IF NOT FRowPrepared THEN
    SelectRow();
    FCapture.Reset();
    IF NOT FPreserveResults THEN
        ResetSubjects();
    END_IF;
    CallSubjects(Enable := FALSE);
    FRowPrepared := TRUE;
ELSE
    CallSubjects(Enable := TRUE);
    CheckResults();
    FObservationReady := TRUE;
END_IF;
END_METHOD

{region 'Documentation'}
(*!
<summary>Requests fresh subject results before the next disabled call.</summary>
*)
{endregion}
METHOD PRIVATE ResetSubjects
FInRangeSubject.Reset();
FNotInRangeSubject.Reset();
END_METHOD

{region 'Documentation'}
(*!
<summary>Selects literal expectations; only named escalation rows retain preceding subject results.</summary>
*)
{endregion}
METHOD PRIVATE SelectRow
FPreserveResults := FALSE;
CASE FRow OF
    LowerEndpoint:
        FActual := ULINT#9223372036854775807;
        FLower := ULINT#9223372036854775807;
        FUpper := ULINT#9223372036854775809;
        FExpectedInRangeResult := E_Result.Passed;
        FExpectedNotInRangeResult := E_Result.Failed;
        FExpectedFindings := 1;
    Interior:
        FActual := ULINT#9223372036854775808;
        FLower := ULINT#9223372036854775807;
        FUpper := ULINT#9223372036854775809;
        FExpectedInRangeResult := E_Result.Passed;
        FExpectedNotInRangeResult := E_Result.Failed;
        FExpectedFindings := 1;
    UpperEndpoint:
        FActual := ULINT#9223372036854775809;
        FLower := ULINT#9223372036854775807;
        FUpper := ULINT#9223372036854775809;
        FExpectedInRangeResult := E_Result.Passed;
        FExpectedNotInRangeResult := E_Result.Failed;
        FExpectedFindings := 1;
    BelowRange:
        FActual := ULINT#9223372036854775806;
        FLower := ULINT#9223372036854775807;
        FUpper := ULINT#9223372036854775809;
        FExpectedInRangeResult := E_Result.Failed;
        FExpectedNotInRangeResult := E_Result.Passed;
        FExpectedFindings := 1;
    AboveRange:
        FActual := ULINT#9223372036854775810;
        FLower := ULINT#9223372036854775807;
        FUpper := ULINT#9223372036854775809;
        FExpectedInRangeResult := E_Result.Failed;
        FExpectedNotInRangeResult := E_Result.Passed;
        FExpectedFindings := 1;
    EqualBounds:
        FActual := ULINT#9223372036854775808;
        FLower := ULINT#9223372036854775808;
        FUpper := ULINT#9223372036854775808;
        FExpectedInRangeResult := E_Result.Passed;
        FExpectedNotInRangeResult := E_Result.Failed;
        FExpectedFindings := 1;
    ReversedBounds:
        FActual := ULINT#9223372036854775808;
        FLower := ULINT#9223372036854775809;
        FUpper := ULINT#9223372036854775807;
        FExpectedInRangeResult := E_Result.Error;
        FExpectedNotInRangeResult := E_Result.Error;
        FExpectedFindings := 2;
    MinimumEndpoint:
        FActual := LowestValue;
        FLower := LowestValue;
        FUpper := HighestValue;
        FExpectedInRangeResult := E_Result.Passed;
        FExpectedNotInRangeResult := E_Result.Failed;
        FExpectedFindings := 1;
    MaximumEndpoint:
        FActual := HighestValue;
        FLower := LowestValue;
        FUpper := HighestValue;
        FExpectedInRangeResult := E_Result.Passed;
        FExpectedNotInRangeResult := E_Result.Failed;
        FExpectedFindings := 1;
    FailureBeforeInvalid:
        FActual := ULINT#9223372036854775810;
        FLower := ULINT#9223372036854775807;
        FUpper := ULINT#9223372036854775809;
        FExpectedInRangeResult := E_Result.Failed;
        FExpectedNotInRangeResult := E_Result.Passed;
        FExpectedFindings := 1;
    InvalidAfterFailure:
        FActual := ULINT#9223372036854775808;
        FLower := ULINT#9223372036854775809;
        FUpper := ULINT#9223372036854775807;
        FExpectedInRangeResult := E_Result.Error;
        FExpectedNotInRangeResult := E_Result.Error;
        FExpectedFindings := 2;
        FPreserveResults := TRUE;
ELSE
    Error(Message := 'Unknown comparison test row.');
END_CASE;
END_METHOD

END_FUNCTION_BLOCK

// ---- SelfTests/TestCases/TestSuite_AssertionComparisons/Test_AssertionDurationComparisons.TcPOU
{region 'Documentation'}
(*!
<summary>Checks duration operators at millisecond boundaries and LTIME nanosecond resolution.</summary>
<description>
Named rows separate independent comparisons by a disabled reset call.
Only explicitly marked escalation rows retain the preceding subject result.
Outer Assertions latch every observation before advancing to the next row.
Intentional findings remain in the local capture; no production algorithm is copied.
</description>
*)
{endregion}
FUNCTION_BLOCK Test_AssertionDurationComparisons EXTENDS TestCaseBase
VAR
    FEqualSubject : AssertEqual_Time;
    FNotEqualSubject : AssertNotEqual_Time;
    FEarlierThanSubject : AssertEarlierThan_Time;
    FLaterThanSubject : AssertLaterThan_Time;
    FInTimespanSubject : AssertInTimespan_Time;
    FNotInTimespanSubject : AssertNotInTimespan_Time;
    FEqualLTimeSubject : AssertEqual_LTime;
    FActual : TIME;
    FReference : TIME;
    FStart : TIME;
    FEnd : TIME;
    FActualLong : LTIME;
    FReferenceLong : LTIME;
    FExpectedEqualResult : E_Result;
    FExpectedNotEqualResult : E_Result;
    FExpectedEarlierThanResult : E_Result;
    FExpectedLaterThanResult : E_Result;
    FExpectedInTimespanResult : E_Result;
    FExpectedNotInTimespanResult : E_Result;
    FExpectedEqualLTimeResult : E_Result;
    FExpectedFindings : UDINT;
    FCapture : EventBuffer;
    FEvents : ARRAY[1..CaptureLength] OF ST_Event;
    FCaptureFifo : ST_FifoStatus;
    FCaptureStatus : ST_EventBufferStatus;
    FRow : UINT;
    FRowPrepared : BOOL;
    FPreserveResults : BOOL;
    FObservationReady : BOOL;
    FChecked : BOOL;
    FSetupValid : BOOL;
END_VAR
VAR
    FEqualResult : AssertTrue;
    FEqualResultMatches : BOOL;
    FNotEqualResult : AssertTrue;
    FNotEqualResultMatches : BOOL;
    FEarlierThanResult : AssertTrue;
    FEarlierThanResultMatches : BOOL;
    FLaterThanResult : AssertTrue;
    FLaterThanResultMatches : BOOL;
    FInTimespanResult : AssertTrue;
    FInTimespanResultMatches : BOOL;
    FNotInTimespanResult : AssertTrue;
    FNotInTimespanResultMatches : BOOL;
    FEqualLTimeResult : AssertTrue;
    FEqualLTimeResultMatches : BOOL;
    FCaptureIntegrity : AssertTrue;
    FCaptureIntegrityMatches : BOOL;
END_VAR
VAR CONSTANT
    CaptureLength : UINT := 8;
    Below : UINT := 1;
    Equal : UINT := 2;
    Above : UINT := 3;
    Outside : UINT := 4;
    EqualBounds : UINT := 5;
    ReversedBounds : UINT := 6;
    LastRow : UINT := ReversedBounds;

END_VAR

SUPER^();

{region 'Documentation'}
(*!
<summary>Collects only outer checking Assertions, never intentional subject findings.</summary>
*)
{endregion}
METHOD PROTECTED AggregateResults
VAR_INPUT
    Aggregator : I_ResultAggregator; //! Borrowed result sink owned by the outer Test Case; add this test's checking Assertions without resetting or retaining the sink.
END_VAR
Aggregator.AddProvider(Provider := FEqualResult);
Aggregator.AddProvider(Provider := FNotEqualResult);
Aggregator.AddProvider(Provider := FEarlierThanResult);
Aggregator.AddProvider(Provider := FLaterThanResult);
Aggregator.AddProvider(Provider := FInTimespanResult);
Aggregator.AddProvider(Provider := FNotInTimespanResult);
Aggregator.AddProvider(Provider := FEqualLTimeResult);
Aggregator.AddProvider(Provider := FCaptureIntegrity);
END_METHOD

{region 'Documentation'}
(*!
<summary>Calls each inherited production Assertion once using the selected row.</summary>
*)
{endregion}
METHOD PRIVATE CallSubjects
VAR_INPUT
    Enable : BOOL; //! Observation-enable input forwarded to the controlled Assertion subjects for this call.
END_VAR
FEqualSubject(Enable := Enable,
    State := E_State.Running,
    IN := FActual,
    Expected := FReference);
FNotEqualSubject(Enable := Enable,
    State := E_State.Running,
    IN := FActual,
    Expected := FReference);
FEarlierThanSubject(Enable := Enable,
    State := E_State.Running,
    IN := FActual,
    Maximum := FReference);
FLaterThanSubject(Enable := Enable,
    State := E_State.Running,
    IN := FActual,
    Minimum := FReference);
FInTimespanSubject(Enable := Enable,
    State := E_State.Running,
    IN := FActual,
    StartTime := FStart,
    EndTime := FEnd);
FNotInTimespanSubject(Enable := Enable,
    State := E_State.Running,
    IN := FActual,
    StartTime := FStart,
    EndTime := FEnd);
FEqualLTimeSubject(Enable := Enable,
    State := E_State.Running,
    IN := FActualLong,
    Expected := FReferenceLong);
END_METHOD

{region 'Documentation'}
(*!
<summary>Extends base validation with subject and checking-Assertion setup.</summary>
*)
{endregion}
METHOD PROTECTED CheckInitialization : BOOL //! TRUE when the inherited initialization check and this concrete fixture check both accept the setup.
CheckInitialization := SUPER^.CheckInitialization();
IF NOT CheckInitialization THEN
    RETURN;
END_IF;

CheckInitialization := FSetupValid
    AND FEqualResult.IsInitialized
    AND FNotEqualResult.IsInitialized
    AND FEarlierThanResult.IsInitialized
    AND FLaterThanResult.IsInitialized
    AND FInTimespanResult.IsInitialized
    AND FNotInTimespanResult.IsInitialized
    AND FEqualLTimeResult.IsInitialized
    AND FCaptureIntegrity.IsInitialized;
IF NOT CheckInitialization THEN
    EventPublisher.PublishEvent(Event := CreateFrameworkEvent(Name := Name,
        ResourceName := '',
        State := State,
        Severity := E_EventSeverity.Error,
        Message := 'Comparison selftest setup failed.'));
END_IF;
END_METHOD

{region 'Documentation'}
(*!
<summary>Checks results and isolated findings against explicit expectations.</summary>
*)
{endregion}
METHOD PRIVATE CheckResults
FEqualResultMatches := FEqualSubject.Result = FExpectedEqualResult;
FNotEqualResultMatches := FNotEqualSubject.Result = FExpectedNotEqualResult;
FEarlierThanResultMatches := FEarlierThanSubject.Result = FExpectedEarlierThanResult;
FLaterThanResultMatches := FLaterThanSubject.Result = FExpectedLaterThanResult;
FInTimespanResultMatches := FInTimespanSubject.Result = FExpectedInTimespanResult;
FNotInTimespanResultMatches := FNotInTimespanSubject.Result = FExpectedNotInTimespanResult;
FEqualLTimeResultMatches := FEqualLTimeSubject.Result = FExpectedEqualLTimeResult;
FCaptureIntegrityMatches := (FCaptureStatus.SequenceId = FExpectedFindings)
    AND (FCaptureStatus.LostEventCount = 0);
END_METHOD

{region 'Documentation'}
(*!
<summary>Configures checking Assertions; subject actions remain in the test script.</summary>
*)
{endregion}
METHOD PROTECTED Configure
VAR
    Initialized : BOOL;
END_VAR
FPreparationStateCount := 0;
FTestStateCount := 1;
FEqualResult.Initialize(Parent := THIS^,
    AssertionName := 'EqualResult');
FNotEqualResult.Initialize(Parent := THIS^,
    AssertionName := 'NotEqualResult');
FEarlierThanResult.Initialize(Parent := THIS^,
    AssertionName := 'EarlierThanResult');
FLaterThanResult.Initialize(Parent := THIS^,
    AssertionName := 'LaterThanResult');
FInTimespanResult.Initialize(Parent := THIS^,
    AssertionName := 'InTimespanResult');
FNotInTimespanResult.Initialize(Parent := THIS^,
    AssertionName := 'NotInTimespanResult');
FEqualLTimeResult.Initialize(Parent := THIS^,
    AssertionName := 'EqualLTimeResult');
FCaptureIntegrity.Initialize(Parent := THIS^,
    AssertionName := 'CaptureIntegrity');
FSetupValid := FCapture.Initialize(Buffer := FEvents,
    FifoControl := FCaptureFifo,
    Status := FCaptureStatus);
FEqualSubject.BindPublisher(Publisher := FCapture);
Initialized := FEqualSubject.Initialize(Parent := THIS^,
    AssertionName := 'EqualSubject');
FSetupValid := FSetupValid AND Initialized;
FNotEqualSubject.BindPublisher(Publisher := FCapture);
Initialized := FNotEqualSubject.Initialize(Parent := THIS^,
    AssertionName := 'NotEqualSubject');
FSetupValid := FSetupValid AND Initialized;
FEarlierThanSubject.BindPublisher(Publisher := FCapture);
Initialized := FEarlierThanSubject.Initialize(Parent := THIS^,
    AssertionName := 'EarlierThanSubject');
FSetupValid := FSetupValid AND Initialized;
FLaterThanSubject.BindPublisher(Publisher := FCapture);
Initialized := FLaterThanSubject.Initialize(Parent := THIS^,
    AssertionName := 'LaterThanSubject');
FSetupValid := FSetupValid AND Initialized;
FInTimespanSubject.BindPublisher(Publisher := FCapture);
Initialized := FInTimespanSubject.Initialize(Parent := THIS^,
    AssertionName := 'InTimespanSubject');
FSetupValid := FSetupValid AND Initialized;
FNotInTimespanSubject.BindPublisher(Publisher := FCapture);
Initialized := FNotInTimespanSubject.Initialize(Parent := THIS^,
    AssertionName := 'NotInTimespanSubject');
FSetupValid := FSetupValid AND Initialized;
FEqualLTimeSubject.BindPublisher(Publisher := FCapture);
Initialized := FEqualLTimeSubject.Initialize(Parent := THIS^,
    AssertionName := 'EqualLTimeSubject');
FSetupValid := FSetupValid AND Initialized;
END_METHOD

{region 'Documentation'}
(*!
<summary>Completes abort without asynchronous resources.</summary>
*)
{endregion}
METHOD PROTECTED ProcessAbort
VAR_INPUT
    Enable : BOOL; //! Phase permission supplied by the owning Test Case; FALSE does not authorize progression, while observation may continue.
END_VAR
IF Enable THEN
    CompleteAbort();
END_IF;
END_METHOD

{region 'Documentation'}
(*!
<summary>Latches checked observations before the next script step may proceed.</summary>
*)
{endregion}
METHOD PROTECTED ProcessAssertions
VAR_INPUT
    Enable : BOOL; //! Phase permission supplied by the owning Test Case; FALSE does not authorize progression, while observation may continue.
END_VAR
VAR
    Evaluate : BOOL;
END_VAR
Evaluate := Enable AND FObservationReady;
FEqualResult(Enable := Evaluate,
    State := State,
    IN := FEqualResultMatches);
FNotEqualResult(Enable := Evaluate,
    State := State,
    IN := FNotEqualResultMatches);
FEarlierThanResult(Enable := Evaluate,
    State := State,
    IN := FEarlierThanResultMatches);
FLaterThanResult(Enable := Evaluate,
    State := State,
    IN := FLaterThanResultMatches);
FInTimespanResult(Enable := Evaluate,
    State := State,
    IN := FInTimespanResultMatches);
FNotInTimespanResult(Enable := Evaluate,
    State := State,
    IN := FNotInTimespanResultMatches);
FEqualLTimeResult(Enable := Evaluate,
    State := State,
    IN := FEqualLTimeResultMatches);
FCaptureIntegrity(Enable := Evaluate,
    State := State,
    IN := FCaptureIntegrityMatches);
IF Evaluate THEN
    FChecked := TRUE;
END_IF;
END_METHOD

{region 'Documentation'}
(*!
<summary>No Preparation phase is required.</summary>
*)
{endregion}
METHOD PROTECTED ProcessPreparations
VAR_INPUT
    // SA0033: Required hook; this test has no Preparation phase.
    {attribute 'analysis' := '-33'}
    Enable : BOOL; //! Phase permission supplied by the owning Test Case; FALSE does not authorize progression, while observation may continue.
END_VAR
END_METHOD

{region 'Documentation'}
(*!
<summary>Restarts the script and resets the checking Assertions.</summary>
*)
{endregion}
METHOD PROTECTED ProcessReset
FRow := Below;
FRowPrepared := FALSE;
FChecked := FALSE;
FObservationReady := FALSE;
FEqualResult.Reset();
FEqualResultMatches := TRUE;
FNotEqualResult.Reset();
FNotEqualResultMatches := TRUE;
FEarlierThanResult.Reset();
FEarlierThanResultMatches := TRUE;
FLaterThanResult.Reset();
FLaterThanResultMatches := TRUE;
FInTimespanResult.Reset();
FInTimespanResultMatches := TRUE;
FNotInTimespanResult.Reset();
FNotInTimespanResultMatches := TRUE;
FEqualLTimeResult.Reset();
FEqualLTimeResultMatches := TRUE;
FCaptureIntegrity.Reset();
FCaptureIntegrityMatches := TRUE;
CompleteReset();
END_METHOD

{region 'Documentation'}
(*!
<summary>Advances one bounded script step per active PLC cycle.</summary>
*)
{endregion}
METHOD PROTECTED ProcessTests
VAR_INPUT
    Enable : BOOL; //! Phase permission supplied by the owning Test Case; FALSE does not authorize progression, while observation may continue.
END_VAR
IF NOT Enable THEN
    RETURN;
END_IF;

IF FChecked THEN
    FChecked := FALSE;
    FObservationReady := FALSE;
    IF FRow = LastRow THEN
        CompleteTests();
        RETURN;
    END_IF;
    FRow := FRow + 1;
    FRowPrepared := FALSE;
END_IF;

IF NOT FRowPrepared THEN
    SelectRow();
    FCapture.Reset();
    IF NOT FPreserveResults THEN
        ResetSubjects();
    END_IF;
    CallSubjects(Enable := FALSE);
    FRowPrepared := TRUE;
ELSE
    CallSubjects(Enable := TRUE);
    CheckResults();
    FObservationReady := TRUE;
END_IF;
END_METHOD

{region 'Documentation'}
(*!
<summary>Requests fresh subject results before the next disabled call.</summary>
*)
{endregion}
METHOD PRIVATE ResetSubjects
FEqualSubject.Reset();
FNotEqualSubject.Reset();
FEarlierThanSubject.Reset();
FLaterThanSubject.Reset();
FInTimespanSubject.Reset();
FNotInTimespanSubject.Reset();
FEqualLTimeSubject.Reset();
END_METHOD

{region 'Documentation'}
(*!
<summary>Selects literal expectations; only named escalation rows retain preceding subject results.</summary>
*)
{endregion}
METHOD PRIVATE SelectRow
FPreserveResults := FALSE;
CASE FRow OF
    Below:
        FActual := T#0ms;
        FReference := T#1ms;
        FStart := T#0ms;
        FEnd := T#2ms;
        FActualLong := LTIME#0ns;
        FReferenceLong := LTIME#1ns;
        FExpectedEqualResult := E_Result.Failed;
        FExpectedNotEqualResult := E_Result.Passed;
        FExpectedEarlierThanResult := E_Result.Passed;
        FExpectedLaterThanResult := E_Result.Failed;
        FExpectedInTimespanResult := E_Result.Passed;
        FExpectedNotInTimespanResult := E_Result.Failed;
        FExpectedEqualLTimeResult := E_Result.Failed;
        FExpectedFindings := 4;
    Equal:
        FActual := T#1ms;
        FReference := T#1ms;
        FStart := T#0ms;
        FEnd := T#2ms;
        FActualLong := LTIME#1ns;
        FReferenceLong := LTIME#1ns;
        FExpectedEqualResult := E_Result.Passed;
        FExpectedNotEqualResult := E_Result.Failed;
        FExpectedEarlierThanResult := E_Result.Failed;
        FExpectedLaterThanResult := E_Result.Failed;
        FExpectedInTimespanResult := E_Result.Passed;
        FExpectedNotInTimespanResult := E_Result.Failed;
        FExpectedEqualLTimeResult := E_Result.Passed;
        FExpectedFindings := 4;
    Above:
        FActual := T#2ms;
        FReference := T#1ms;
        FStart := T#0ms;
        FEnd := T#2ms;
        FActualLong := LTIME#2ns;
        FReferenceLong := LTIME#1ns;
        FExpectedEqualResult := E_Result.Failed;
        FExpectedNotEqualResult := E_Result.Passed;
        FExpectedEarlierThanResult := E_Result.Failed;
        FExpectedLaterThanResult := E_Result.Passed;
        FExpectedInTimespanResult := E_Result.Passed;
        FExpectedNotInTimespanResult := E_Result.Failed;
        FExpectedEqualLTimeResult := E_Result.Failed;
        FExpectedFindings := 4;
    Outside:
        FActual := T#3ms;
        FReference := T#1ms;
        FStart := T#0ms;
        FEnd := T#2ms;
        FActualLong := LTIME#0ns;
        FReferenceLong := LTIME#1ns;
        FExpectedEqualResult := E_Result.Failed;
        FExpectedNotEqualResult := E_Result.Passed;
        FExpectedEarlierThanResult := E_Result.Failed;
        FExpectedLaterThanResult := E_Result.Passed;
        FExpectedInTimespanResult := E_Result.Failed;
        FExpectedNotInTimespanResult := E_Result.Passed;
        FExpectedEqualLTimeResult := E_Result.Failed;
        FExpectedFindings := 4;
    EqualBounds:
        FActual := T#1ms;
        FReference := T#1ms;
        FStart := T#1ms;
        FEnd := T#1ms;
        FActualLong := LTIME#1ns;
        FReferenceLong := LTIME#1ns;
        FExpectedEqualResult := E_Result.Passed;
        FExpectedNotEqualResult := E_Result.Failed;
        FExpectedEarlierThanResult := E_Result.Failed;
        FExpectedLaterThanResult := E_Result.Failed;
        FExpectedInTimespanResult := E_Result.Passed;
        FExpectedNotInTimespanResult := E_Result.Failed;
        FExpectedEqualLTimeResult := E_Result.Passed;
        FExpectedFindings := 4;
    ReversedBounds:
        FActual := T#1ms;
        FReference := T#1ms;
        FStart := T#2ms;
        FEnd := T#0ms;
        FActualLong := LTIME#1ns;
        FReferenceLong := LTIME#1ns;
        FExpectedEqualResult := E_Result.Passed;
        FExpectedNotEqualResult := E_Result.Failed;
        FExpectedEarlierThanResult := E_Result.Failed;
        FExpectedLaterThanResult := E_Result.Failed;
        FExpectedInTimespanResult := E_Result.Error;
        FExpectedNotInTimespanResult := E_Result.Error;
        FExpectedEqualLTimeResult := E_Result.Passed;
        FExpectedFindings := 5;
ELSE
    Error(Message := 'Unknown comparison test row.');
END_CASE;
END_METHOD

END_FUNCTION_BLOCK

// ---- Framework/Assertions/POU/BasicTypes/LTime/AssertEqual_LTime.TcPOU
{region 'Documentation'}
(*!
<summary>Checks equality with the expected LTIME value.</summary>
*)
{endregion}
FUNCTION_BLOCK AssertEqual_LTime EXTENDS AssertionBase
VAR_INPUT
    IN : LTIME; //! Actual value checked or observed by this Assertion.
    Expected : LTIME; //! Reference value for comparison with IN.
END_VAR

SUPER^();

{region 'Documentation'}
(*!
<summary>Evaluate the typed duration relation and report higher-priority errors first.</summary>
*)
{endregion}
METHOD PROTECTED Assert
VAR
    Message : STRING(GVL_Constants.MessageLength);
    ExpectedText : STRING(GVL_Constants.AssertionValueLength);
    ActualText : STRING(GVL_Constants.AssertionValueLength);
END_VAR
IF NOT EvaluationActive THEN
    RETURN;
END_IF;

IF Result = E_Result.Error THEN
    RETURN;
END_IF;

IF Result = E_Result.Failed THEN
    RETURN;
END_IF;

IF IN <> Expected THEN
    ExpectedText := LTIME_TO_STRING(Expected);
    ActualText := LTIME_TO_STRING(IN);
    Message := CONCAT('Assertion failed: values are not equal. Expected = ',
        ExpectedText);
    Message := CONCAT(Message, ', Actual = ');
    Message := CONCAT(Message, ActualText);
    Message := CONCAT(Message, '.');
    Fail(Message := Message);
    RETURN;
END_IF;

Pass();
END_METHOD

END_FUNCTION_BLOCK

// ---- SelfTests/TestCases/TestSuite_AssertionComparisons/Test_AssertionDateNormalization.TcPOU
{region 'Documentation'}
(*!
<summary>Checks calendar-day identity and range bounds despite hidden time-of-day components.</summary>
<description>
Named rows separate independent comparisons by a disabled reset call.
Only explicitly marked escalation rows retain the preceding subject result.
Outer Assertions latch every observation before advancing to the next row.
Intentional findings remain in the local capture; no production algorithm is copied.
</description>
*)
{endregion}
FUNCTION_BLOCK Test_AssertionDateNormalization EXTENDS TestCaseBase
VAR
    FEqualSubject : AssertEqual_Date;
    FInTimespanSubject : AssertInTimespan_Date;
    FNotInTimespanSubject : AssertNotInTimespan_Date;
    FActual : DATE;
    FReference : DATE;
    FStart : DATE;
    FEnd : DATE;
    FExpectedEqualResult : E_Result;
    FExpectedInTimespanResult : E_Result;
    FExpectedNotInTimespanResult : E_Result;
    FExpectedFindings : UDINT;
    FCapture : EventBuffer;
    FEvents : ARRAY[1..CaptureLength] OF ST_Event;
    FCaptureFifo : ST_FifoStatus;
    FCaptureStatus : ST_EventBufferStatus;
    FRow : UINT;
    FRowPrepared : BOOL;
    FPreserveResults : BOOL;
    FObservationReady : BOOL;
    FChecked : BOOL;
    FSetupValid : BOOL;
END_VAR
VAR
    FEqualResult : AssertTrue;
    FEqualResultMatches : BOOL;
    FInTimespanResult : AssertTrue;
    FInTimespanResultMatches : BOOL;
    FNotInTimespanResult : AssertTrue;
    FNotInTimespanResultMatches : BOOL;
    FCaptureIntegrity : AssertTrue;
    FCaptureIntegrityMatches : BOOL;
END_VAR
VAR CONSTANT
    CaptureLength : UINT := 8;
    SameDay : UINT := 1;
    NextDay : UINT := 2;
    NormalizedEqualBounds : UINT := 3;
    ReversedDays : UINT := 4;
    LastRow : UINT := ReversedDays;

END_VAR

SUPER^();

{region 'Documentation'}
(*!
<summary>Collects only outer checking Assertions, never intentional subject findings.</summary>
*)
{endregion}
METHOD PROTECTED AggregateResults
VAR_INPUT
    Aggregator : I_ResultAggregator; //! Borrowed result sink owned by the outer Test Case; add this test's checking Assertions without resetting or retaining the sink.
END_VAR
Aggregator.AddProvider(Provider := FEqualResult);
Aggregator.AddProvider(Provider := FInTimespanResult);
Aggregator.AddProvider(Provider := FNotInTimespanResult);
Aggregator.AddProvider(Provider := FCaptureIntegrity);
END_METHOD

{region 'Documentation'}
(*!
<summary>Calls each inherited production Assertion once using the selected row.</summary>
*)
{endregion}
METHOD PRIVATE CallSubjects
VAR_INPUT
    Enable : BOOL; //! Observation-enable input forwarded to the controlled Assertion subjects for this call.
END_VAR
FEqualSubject(Enable := Enable,
    State := E_State.Running,
    IN := FActual,
    Expected := FReference);
FInTimespanSubject(Enable := Enable,
    State := E_State.Running,
    IN := FActual,
    StartTime := FStart,
    EndTime := FEnd);
FNotInTimespanSubject(Enable := Enable,
    State := E_State.Running,
    IN := FActual,
    StartTime := FStart,
    EndTime := FEnd);
END_METHOD

{region 'Documentation'}
(*!
<summary>Extends base validation with subject and checking-Assertion setup.</summary>
*)
{endregion}
METHOD PROTECTED CheckInitialization : BOOL //! TRUE when the inherited initialization check and this concrete fixture check both accept the setup.
CheckInitialization := SUPER^.CheckInitialization();
IF NOT CheckInitialization THEN
    RETURN;
END_IF;

CheckInitialization := FSetupValid
    AND FEqualResult.IsInitialized
    AND FInTimespanResult.IsInitialized
    AND FNotInTimespanResult.IsInitialized
    AND FCaptureIntegrity.IsInitialized;
IF NOT CheckInitialization THEN
    EventPublisher.PublishEvent(Event := CreateFrameworkEvent(Name := Name,
        ResourceName := '',
        State := State,
        Severity := E_EventSeverity.Error,
        Message := 'Comparison selftest setup failed.'));
END_IF;
END_METHOD

{region 'Documentation'}
(*!
<summary>Checks results and isolated findings against explicit expectations.</summary>
*)
{endregion}
METHOD PRIVATE CheckResults
FEqualResultMatches := FEqualSubject.Result = FExpectedEqualResult;
FInTimespanResultMatches := FInTimespanSubject.Result = FExpectedInTimespanResult;
FNotInTimespanResultMatches := FNotInTimespanSubject.Result = FExpectedNotInTimespanResult;
FCaptureIntegrityMatches := (FCaptureStatus.SequenceId = FExpectedFindings)
    AND (FCaptureStatus.LostEventCount = 0);
END_METHOD

{region 'Documentation'}
(*!
<summary>Configures checking Assertions; subject actions remain in the test script.</summary>
*)
{endregion}
METHOD PROTECTED Configure
VAR
    Initialized : BOOL;
END_VAR
FPreparationStateCount := 0;
FTestStateCount := 1;
FEqualResult.Initialize(Parent := THIS^,
    AssertionName := 'EqualResult');
FInTimespanResult.Initialize(Parent := THIS^,
    AssertionName := 'InTimespanResult');
FNotInTimespanResult.Initialize(Parent := THIS^,
    AssertionName := 'NotInTimespanResult');
FCaptureIntegrity.Initialize(Parent := THIS^,
    AssertionName := 'CaptureIntegrity');
FSetupValid := FCapture.Initialize(Buffer := FEvents,
    FifoControl := FCaptureFifo,
    Status := FCaptureStatus);
FEqualSubject.BindPublisher(Publisher := FCapture);
Initialized := FEqualSubject.Initialize(Parent := THIS^,
    AssertionName := 'EqualSubject');
FSetupValid := FSetupValid AND Initialized;
FInTimespanSubject.BindPublisher(Publisher := FCapture);
Initialized := FInTimespanSubject.Initialize(Parent := THIS^,
    AssertionName := 'InTimespanSubject');
FSetupValid := FSetupValid AND Initialized;
FNotInTimespanSubject.BindPublisher(Publisher := FCapture);
Initialized := FNotInTimespanSubject.Initialize(Parent := THIS^,
    AssertionName := 'NotInTimespanSubject');
FSetupValid := FSetupValid AND Initialized;
END_METHOD

{region 'Documentation'}
(*!
<summary>Completes abort without asynchronous resources.</summary>
*)
{endregion}
METHOD PROTECTED ProcessAbort
VAR_INPUT
    Enable : BOOL; //! Phase permission supplied by the owning Test Case; FALSE does not authorize progression, while observation may continue.
END_VAR
IF Enable THEN
    CompleteAbort();
END_IF;
END_METHOD

{region 'Documentation'}
(*!
<summary>Latches checked observations before the next script step may proceed.</summary>
*)
{endregion}
METHOD PROTECTED ProcessAssertions
VAR_INPUT
    Enable : BOOL; //! Phase permission supplied by the owning Test Case; FALSE does not authorize progression, while observation may continue.
END_VAR
VAR
    Evaluate : BOOL;
END_VAR
Evaluate := Enable AND FObservationReady;
FEqualResult(Enable := Evaluate,
    State := State,
    IN := FEqualResultMatches);
FInTimespanResult(Enable := Evaluate,
    State := State,
    IN := FInTimespanResultMatches);
FNotInTimespanResult(Enable := Evaluate,
    State := State,
    IN := FNotInTimespanResultMatches);
FCaptureIntegrity(Enable := Evaluate,
    State := State,
    IN := FCaptureIntegrityMatches);
IF Evaluate THEN
    FChecked := TRUE;
END_IF;
END_METHOD

{region 'Documentation'}
(*!
<summary>No Preparation phase is required.</summary>
*)
{endregion}
METHOD PROTECTED ProcessPreparations
VAR_INPUT
    // SA0033: Required hook; this test has no Preparation phase.
    {attribute 'analysis' := '-33'}
    Enable : BOOL; //! Phase permission supplied by the owning Test Case; FALSE does not authorize progression, while observation may continue.
END_VAR
END_METHOD

{region 'Documentation'}
(*!
<summary>Restarts the script and resets the checking Assertions.</summary>
*)
{endregion}
METHOD PROTECTED ProcessReset
FRow := SameDay;
FRowPrepared := FALSE;
FChecked := FALSE;
FObservationReady := FALSE;
FEqualResult.Reset();
FEqualResultMatches := TRUE;
FInTimespanResult.Reset();
FInTimespanResultMatches := TRUE;
FNotInTimespanResult.Reset();
FNotInTimespanResultMatches := TRUE;
FCaptureIntegrity.Reset();
FCaptureIntegrityMatches := TRUE;
CompleteReset();
END_METHOD

{region 'Documentation'}
(*!
<summary>Advances one bounded script step per active PLC cycle.</summary>
*)
{endregion}
METHOD PROTECTED ProcessTests
VAR_INPUT
    Enable : BOOL; //! Phase permission supplied by the owning Test Case; FALSE does not authorize progression, while observation may continue.
END_VAR
IF NOT Enable THEN
    RETURN;
END_IF;

IF FChecked THEN
    FChecked := FALSE;
    FObservationReady := FALSE;
    IF FRow = LastRow THEN
        CompleteTests();
        RETURN;
    END_IF;
    FRow := FRow + 1;
    FRowPrepared := FALSE;
END_IF;

IF NOT FRowPrepared THEN
    SelectRow();
    FCapture.Reset();
    IF NOT FPreserveResults THEN
        ResetSubjects();
    END_IF;
    CallSubjects(Enable := FALSE);
    FRowPrepared := TRUE;
ELSE
    CallSubjects(Enable := TRUE);
    CheckResults();
    FObservationReady := TRUE;
END_IF;
END_METHOD

{region 'Documentation'}
(*!
<summary>Requests fresh subject results before the next disabled call.</summary>
*)
{endregion}
METHOD PRIVATE ResetSubjects
FEqualSubject.Reset();
FInTimespanSubject.Reset();
FNotInTimespanSubject.Reset();
END_METHOD

{region 'Documentation'}
(*!
<summary>Selects literal expectations; only named escalation rows retain preceding subject results.</summary>
*)
{endregion}
METHOD PRIVATE SelectRow
FPreserveResults := FALSE;
CASE FRow OF
    SameDay:
        FActual := UDINT_TO_DATE(UDINT#172799);
        FReference := UDINT_TO_DATE(UDINT#86400);
        FStart := UDINT_TO_DATE(UDINT#86400);
        FEnd := UDINT_TO_DATE(UDINT#172799);
        FExpectedEqualResult := E_Result.Passed;
        FExpectedInTimespanResult := E_Result.Passed;
        FExpectedNotInTimespanResult := E_Result.Failed;
        FExpectedFindings := 1;
    NextDay:
        FActual := UDINT_TO_DATE(UDINT#172800);
        FReference := UDINT_TO_DATE(UDINT#86400);
        FStart := UDINT_TO_DATE(UDINT#86400);
        FEnd := UDINT_TO_DATE(UDINT#172799);
        FExpectedEqualResult := E_Result.Failed;
        FExpectedInTimespanResult := E_Result.Failed;
        FExpectedNotInTimespanResult := E_Result.Passed;
        FExpectedFindings := 2;
    NormalizedEqualBounds:
        FActual := UDINT_TO_DATE(UDINT#86400);
        FReference := UDINT_TO_DATE(UDINT#172799);
        FStart := UDINT_TO_DATE(UDINT#172799);
        FEnd := UDINT_TO_DATE(UDINT#86400);
        FExpectedEqualResult := E_Result.Passed;
        FExpectedInTimespanResult := E_Result.Passed;
        FExpectedNotInTimespanResult := E_Result.Failed;
        FExpectedFindings := 1;
    ReversedDays:
        FActual := UDINT_TO_DATE(UDINT#86400);
        FReference := UDINT_TO_DATE(UDINT#86400);
        FStart := UDINT_TO_DATE(UDINT#172800);
        FEnd := UDINT_TO_DATE(UDINT#86400);
        FExpectedEqualResult := E_Result.Passed;
        FExpectedInTimespanResult := E_Result.Error;
        FExpectedNotInTimespanResult := E_Result.Error;
        FExpectedFindings := 2;
ELSE
    Error(Message := 'Unknown comparison test row.');
END_CASE;
END_METHOD

END_FUNCTION_BLOCK

// ---- Framework/Assertions/POU/BasicTypes/Date/AssertEqual_Date.TcPOU
{region 'Documentation'}
(*!
<summary>Checks equality with the expected DATE value.</summary>
<description>

Compares calendar days only; hidden time-of-day components are ignored.

</description>
*)
{endregion}
FUNCTION_BLOCK AssertEqual_Date EXTENDS AssertionBase
VAR_INPUT
    IN : DATE; //! Actual value checked or observed by this Assertion.
    Expected : DATE; //! Reference value for comparison with IN.
END_VAR

SUPER^();

{region 'Documentation'}
(*!
<summary>Evaluate the typed temporal relation and report higher-priority errors first.</summary>
*)
{endregion}
METHOD PROTECTED Assert
VAR
    Message : STRING(GVL_Constants.MessageLength);
    ExpectedText : STRING(GVL_Constants.AssertionValueLength);
    ActualText : STRING(GVL_Constants.AssertionValueLength);
END_VAR
IF NOT EvaluationActive THEN
    RETURN;
END_IF;

IF Result = E_Result.Error THEN
    RETURN;
END_IF;

IF Result = E_Result.Failed THEN
    RETURN;
END_IF;

IF DateToDayNumber(Value := IN) <> DateToDayNumber(Value := Expected) THEN
    ExpectedText := DATE_TO_STRING(Expected);
    ActualText := DATE_TO_STRING(IN);
    Message := CONCAT('Assertion failed: values are not equal. Expected = ',
        ExpectedText);
    Message := CONCAT(Message, ', Actual = ');
    Message := CONCAT(Message, ActualText);
    Message := CONCAT(Message, '.');
    Fail(Message := Message);
    RETURN;
END_IF;

Pass();
END_METHOD

END_FUNCTION_BLOCK

// ---- Framework/Assertions/POU/Utilities/DateToDayNumber.TcPOU
{region 'Documentation'}
(*!
<summary>Returns whole calendar days since 1970-01-01; ignores any time-of-day remainder.</summary>
*)
{endregion}
FUNCTION INTERNAL DateToDayNumber : UDINT //! Whole days since 1970-01-01.
VAR_INPUT
    Value : DATE; //! Calendar date; any stored time-of-day remainder is ignored.
END_VAR
VAR CONSTANT
    SecondsPerDay : UDINT := 86400;
END_VAR

DateToDayNumber := DATE_TO_UDINT(Value) / SecondsPerDay;

END_FUNCTION

// ---- Framework/Assertions/POU/BasicTypes/Date/AssertInTimespan_Date.TcPOU
{region 'Documentation'}
(*!
<summary>Check that IN is inside the inclusive StartTime..EndTime interval.</summary>
<description>

StartTime &gt; EndTime reports Error during active evaluation; equal bounds are
valid.

Compares calendar days only; hidden time-of-day components are ignored.

</description>
*)
{endregion}
FUNCTION_BLOCK AssertInTimespan_Date EXTENDS AssertionBase
VAR_INPUT
    IN : DATE; //! Actual value checked or observed by this Assertion.
    StartTime : DATE; //! Inclusive start of the time span; must not exceed EndTime.
    EndTime : DATE; //! Inclusive end of the time span; must not precede StartTime.
END_VAR

SUPER^();

{region 'Documentation'}
(*!
<summary>Evaluate the typed temporal relation and report higher-priority errors first.</summary>
*)
{endregion}
METHOD PROTECTED Assert
VAR
    Message : STRING(GVL_Constants.MessageLength);
    StartTimeText : STRING(GVL_Constants.AssertionValueLength);
    EndTimeText : STRING(GVL_Constants.AssertionValueLength);
    ActualText : STRING(GVL_Constants.AssertionValueLength);
END_VAR
IF NOT EvaluationActive THEN
    RETURN;
END_IF;

IF Result = E_Result.Error THEN
    RETURN;
END_IF;

IF DateToDayNumber(Value := StartTime) > DateToDayNumber(Value := EndTime) THEN
    StartTimeText := DATE_TO_STRING(StartTime);
    EndTimeText := DATE_TO_STRING(EndTime);
    Message := CONCAT('Assertion error: start time exceeds end time. StartTime = ',
        StartTimeText);
    Message := CONCAT(Message, ', EndTime = ');
    Message := CONCAT(Message, EndTimeText);
    Message := CONCAT(Message, '.');
    Error(Message := Message);
    RETURN;
END_IF;

IF Result = E_Result.Failed THEN
    RETURN;
END_IF;

IF (DateToDayNumber(Value := IN) < DateToDayNumber(Value := StartTime))
    OR (DateToDayNumber(Value := IN) > DateToDayNumber(Value := EndTime)) THEN
    StartTimeText := DATE_TO_STRING(StartTime);
    EndTimeText := DATE_TO_STRING(EndTime);
    ActualText := DATE_TO_STRING(IN);
    Message := CONCAT('Assertion failed: value is outside allowed timespan. StartTime = ',
        StartTimeText);
    Message := CONCAT(Message, ', EndTime = ');
    Message := CONCAT(Message, EndTimeText);
    Message := CONCAT(Message, ', Actual = ');
    Message := CONCAT(Message, ActualText);
    Message := CONCAT(Message, '.');
    Fail(Message := Message);
    RETURN;
END_IF;

Pass();
END_METHOD

END_FUNCTION_BLOCK

// ---- Framework/Assertions/POU/BasicTypes/Date/AssertNotInTimespan_Date.TcPOU
{region 'Documentation'}
(*!
<summary>Check that IN is outside the inclusive StartTime..EndTime interval.</summary>
<description>

StartTime &gt; EndTime reports Error during active evaluation; equal bounds are
valid.

Compares calendar days only; hidden time-of-day components are ignored.

</description>
*)
{endregion}
FUNCTION_BLOCK AssertNotInTimespan_Date EXTENDS AssertionBase
VAR_INPUT
    IN : DATE; //! Actual value checked or observed by this Assertion.
    StartTime : DATE; //! Inclusive start of the time span; must not exceed EndTime.
    EndTime : DATE; //! Inclusive end of the time span; must not precede StartTime.
END_VAR

SUPER^();

{region 'Documentation'}
(*!
<summary>Evaluate the typed temporal relation and report higher-priority errors first.</summary>
*)
{endregion}
METHOD PROTECTED Assert
VAR
    Message : STRING(GVL_Constants.MessageLength);
    StartTimeText : STRING(GVL_Constants.AssertionValueLength);
    EndTimeText : STRING(GVL_Constants.AssertionValueLength);
    ActualText : STRING(GVL_Constants.AssertionValueLength);
END_VAR
IF NOT EvaluationActive THEN
    RETURN;
END_IF;

IF Result = E_Result.Error THEN
    RETURN;
END_IF;

IF DateToDayNumber(Value := StartTime) > DateToDayNumber(Value := EndTime) THEN
    StartTimeText := DATE_TO_STRING(StartTime);
    EndTimeText := DATE_TO_STRING(EndTime);
    Message := CONCAT('Assertion error: start time exceeds end time. StartTime = ',
        StartTimeText);
    Message := CONCAT(Message, ', EndTime = ');
    Message := CONCAT(Message, EndTimeText);
    Message := CONCAT(Message, '.');
    Error(Message := Message);
    RETURN;
END_IF;

IF Result = E_Result.Failed THEN
    RETURN;
END_IF;

IF (DateToDayNumber(Value := IN) >= DateToDayNumber(Value := StartTime))
    AND (DateToDayNumber(Value := IN) <= DateToDayNumber(Value := EndTime)) THEN
    StartTimeText := DATE_TO_STRING(StartTime);
    EndTimeText := DATE_TO_STRING(EndTime);
    ActualText := DATE_TO_STRING(IN);
    Message := CONCAT('Assertion failed: value is inside forbidden timespan. StartTime = ',
        StartTimeText);
    Message := CONCAT(Message, ', EndTime = ');
    Message := CONCAT(Message, EndTimeText);
    Message := CONCAT(Message, ', Actual = ');
    Message := CONCAT(Message, ActualText);
    Message := CONCAT(Message, '.');
    Fail(Message := Message);
    RETURN;
END_IF;

Pass();
END_METHOD

END_FUNCTION_BLOCK

// ---- SelfTests/TestCases/TestSuite_AssertionComparisons/Test_AssertionTODDomain.TcPOU
{region 'Documentation'}
(*!
<summary>Checks all TOD inputs at midnight and the exclusive 24-hour domain limit.</summary>
<description>
Named rows separate independent comparisons by a disabled reset call.
Only explicitly marked escalation rows retain the preceding subject result.
Outer Assertions latch every observation before advancing to the next row.
Intentional findings remain in the local capture; no production algorithm is copied.
</description>
*)
{endregion}
FUNCTION_BLOCK Test_AssertionTODDomain EXTENDS TestCaseBase
VAR
    FEqualSubject : AssertEqual_TOD;
    FInTimespanSubject : AssertInTimespan_TOD;
    FNotInTimespanSubject : AssertNotInTimespan_TOD;
    FActual : TOD;
    FReference : TOD;
    FStart : TOD;
    FEnd : TOD;
    FExpectedEqualResult : E_Result;
    FExpectedInTimespanResult : E_Result;
    FExpectedNotInTimespanResult : E_Result;
    FExpectedFindings : UDINT;
    FCapture : EventBuffer;
    FEvents : ARRAY[1..CaptureLength] OF ST_Event;
    FCaptureFifo : ST_FifoStatus;
    FCaptureStatus : ST_EventBufferStatus;
    FRow : UINT;
    FRowPrepared : BOOL;
    FPreserveResults : BOOL;
    FObservationReady : BOOL;
    FChecked : BOOL;
    FSetupValid : BOOL;
END_VAR
VAR
    FEqualResult : AssertTrue;
    FEqualResultMatches : BOOL;
    FInTimespanResult : AssertTrue;
    FInTimespanResultMatches : BOOL;
    FNotInTimespanResult : AssertTrue;
    FNotInTimespanResultMatches : BOOL;
    FCaptureIntegrity : AssertTrue;
    FCaptureIntegrityMatches : BOOL;
END_VAR
VAR CONSTANT
    CaptureLength : UINT := 8;
    Midnight : UINT := 1;
    LastValidValue : UINT := 2;
    DistinctValid : UINT := 3;
    InvalidInput : UINT := 4;
    InvalidExpected : UINT := 5;
    InvalidStart : UINT := 6;
    InvalidEnd : UINT := 7;
    ReversedValidSpan : UINT := 8;
    LastRow : UINT := ReversedValidSpan;
    Zero : TOD := TOD#00:00:00;
    LastValid : TOD := TOD#23:59:59.999;
    OneDay : TOD := UDINT_TO_TOD(UDINT#86400000);
END_VAR

SUPER^();

{region 'Documentation'}
(*!
<summary>Collects only outer checking Assertions, never intentional subject findings.</summary>
*)
{endregion}
METHOD PROTECTED AggregateResults
VAR_INPUT
    Aggregator : I_ResultAggregator; //! Borrowed result sink owned by the outer Test Case; add this test's checking Assertions without resetting or retaining the sink.
END_VAR
Aggregator.AddProvider(Provider := FEqualResult);
Aggregator.AddProvider(Provider := FInTimespanResult);
Aggregator.AddProvider(Provider := FNotInTimespanResult);
Aggregator.AddProvider(Provider := FCaptureIntegrity);
END_METHOD

{region 'Documentation'}
(*!
<summary>Calls each inherited production Assertion once using the selected row.</summary>
*)
{endregion}
METHOD PRIVATE CallSubjects
VAR_INPUT
    Enable : BOOL; //! Observation-enable input forwarded to the controlled Assertion subjects for this call.
END_VAR
FEqualSubject(Enable := Enable,
    State := E_State.Running,
    IN := FActual,
    Expected := FReference);
FInTimespanSubject(Enable := Enable,
    State := E_State.Running,
    IN := FActual,
    StartTime := FStart,
    EndTime := FEnd);
FNotInTimespanSubject(Enable := Enable,
    State := E_State.Running,
    IN := FActual,
    StartTime := FStart,
    EndTime := FEnd);
END_METHOD

{region 'Documentation'}
(*!
<summary>Extends base validation with subject and checking-Assertion setup.</summary>
*)
{endregion}
METHOD PROTECTED CheckInitialization : BOOL //! TRUE when the inherited initialization check and this concrete fixture check both accept the setup.
CheckInitialization := SUPER^.CheckInitialization();
IF NOT CheckInitialization THEN
    RETURN;
END_IF;

CheckInitialization := FSetupValid
    AND FEqualResult.IsInitialized
    AND FInTimespanResult.IsInitialized
    AND FNotInTimespanResult.IsInitialized
    AND FCaptureIntegrity.IsInitialized;
IF NOT CheckInitialization THEN
    EventPublisher.PublishEvent(Event := CreateFrameworkEvent(Name := Name,
        ResourceName := '',
        State := State,
        Severity := E_EventSeverity.Error,
        Message := 'Comparison selftest setup failed.'));
END_IF;
END_METHOD

{region 'Documentation'}
(*!
<summary>Checks results and isolated findings against explicit expectations.</summary>
*)
{endregion}
METHOD PRIVATE CheckResults
FEqualResultMatches := FEqualSubject.Result = FExpectedEqualResult;
FInTimespanResultMatches := FInTimespanSubject.Result = FExpectedInTimespanResult;
FNotInTimespanResultMatches := FNotInTimespanSubject.Result = FExpectedNotInTimespanResult;
FCaptureIntegrityMatches := (FCaptureStatus.SequenceId = FExpectedFindings)
    AND (FCaptureStatus.LostEventCount = 0);
END_METHOD

{region 'Documentation'}
(*!
<summary>Configures checking Assertions; subject actions remain in the test script.</summary>
*)
{endregion}
METHOD PROTECTED Configure
VAR
    Initialized : BOOL;
END_VAR
FPreparationStateCount := 0;
FTestStateCount := 1;
FEqualResult.Initialize(Parent := THIS^,
    AssertionName := 'EqualResult');
FInTimespanResult.Initialize(Parent := THIS^,
    AssertionName := 'InTimespanResult');
FNotInTimespanResult.Initialize(Parent := THIS^,
    AssertionName := 'NotInTimespanResult');
FCaptureIntegrity.Initialize(Parent := THIS^,
    AssertionName := 'CaptureIntegrity');
FSetupValid := FCapture.Initialize(Buffer := FEvents,
    FifoControl := FCaptureFifo,
    Status := FCaptureStatus);
FEqualSubject.BindPublisher(Publisher := FCapture);
Initialized := FEqualSubject.Initialize(Parent := THIS^,
    AssertionName := 'EqualSubject');
FSetupValid := FSetupValid AND Initialized;
FInTimespanSubject.BindPublisher(Publisher := FCapture);
Initialized := FInTimespanSubject.Initialize(Parent := THIS^,
    AssertionName := 'InTimespanSubject');
FSetupValid := FSetupValid AND Initialized;
FNotInTimespanSubject.BindPublisher(Publisher := FCapture);
Initialized := FNotInTimespanSubject.Initialize(Parent := THIS^,
    AssertionName := 'NotInTimespanSubject');
FSetupValid := FSetupValid AND Initialized;
END_METHOD

{region 'Documentation'}
(*!
<summary>Completes abort without asynchronous resources.</summary>
*)
{endregion}
METHOD PROTECTED ProcessAbort
VAR_INPUT
    Enable : BOOL; //! Phase permission supplied by the owning Test Case; FALSE does not authorize progression, while observation may continue.
END_VAR
IF Enable THEN
    CompleteAbort();
END_IF;
END_METHOD

{region 'Documentation'}
(*!
<summary>Latches checked observations before the next script step may proceed.</summary>
*)
{endregion}
METHOD PROTECTED ProcessAssertions
VAR_INPUT
    Enable : BOOL; //! Phase permission supplied by the owning Test Case; FALSE does not authorize progression, while observation may continue.
END_VAR
VAR
    Evaluate : BOOL;
END_VAR
Evaluate := Enable AND FObservationReady;
FEqualResult(Enable := Evaluate,
    State := State,
    IN := FEqualResultMatches);
FInTimespanResult(Enable := Evaluate,
    State := State,
    IN := FInTimespanResultMatches);
FNotInTimespanResult(Enable := Evaluate,
    State := State,
    IN := FNotInTimespanResultMatches);
FCaptureIntegrity(Enable := Evaluate,
    State := State,
    IN := FCaptureIntegrityMatches);
IF Evaluate THEN
    FChecked := TRUE;
END_IF;
END_METHOD

{region 'Documentation'}
(*!
<summary>No Preparation phase is required.</summary>
*)
{endregion}
METHOD PROTECTED ProcessPreparations
VAR_INPUT
    // SA0033: Required hook; this test has no Preparation phase.
    {attribute 'analysis' := '-33'}
    Enable : BOOL; //! Phase permission supplied by the owning Test Case; FALSE does not authorize progression, while observation may continue.
END_VAR
END_METHOD

{region 'Documentation'}
(*!
<summary>Restarts the script and resets the checking Assertions.</summary>
*)
{endregion}
METHOD PROTECTED ProcessReset
FRow := Midnight;
FRowPrepared := FALSE;
FChecked := FALSE;
FObservationReady := FALSE;
FEqualResult.Reset();
FEqualResultMatches := TRUE;
FInTimespanResult.Reset();
FInTimespanResultMatches := TRUE;
FNotInTimespanResult.Reset();
FNotInTimespanResultMatches := TRUE;
FCaptureIntegrity.Reset();
FCaptureIntegrityMatches := TRUE;
CompleteReset();
END_METHOD

{region 'Documentation'}
(*!
<summary>Advances one bounded script step per active PLC cycle.</summary>
*)
{endregion}
METHOD PROTECTED ProcessTests
VAR_INPUT
    Enable : BOOL; //! Phase permission supplied by the owning Test Case; FALSE does not authorize progression, while observation may continue.
END_VAR
IF NOT Enable THEN
    RETURN;
END_IF;

IF FChecked THEN
    FChecked := FALSE;
    FObservationReady := FALSE;
    IF FRow = LastRow THEN
        CompleteTests();
        RETURN;
    END_IF;
    FRow := FRow + 1;
    FRowPrepared := FALSE;
END_IF;

IF NOT FRowPrepared THEN
    SelectRow();
    FCapture.Reset();
    IF NOT FPreserveResults THEN
        ResetSubjects();
    END_IF;
    CallSubjects(Enable := FALSE);
    FRowPrepared := TRUE;
ELSE
    CallSubjects(Enable := TRUE);
    CheckResults();
    FObservationReady := TRUE;
END_IF;
END_METHOD

{region 'Documentation'}
(*!
<summary>Requests fresh subject results before the next disabled call.</summary>
*)
{endregion}
METHOD PRIVATE ResetSubjects
FEqualSubject.Reset();
FInTimespanSubject.Reset();
FNotInTimespanSubject.Reset();
END_METHOD

{region 'Documentation'}
(*!
<summary>Selects literal expectations; only named escalation rows retain preceding subject results.</summary>
*)
{endregion}
METHOD PRIVATE SelectRow
FPreserveResults := FALSE;
CASE FRow OF
    Midnight:
        FActual := Zero;
        FReference := Zero;
        FStart := Zero;
        FEnd := LastValid;
        FExpectedEqualResult := E_Result.Passed;
        FExpectedInTimespanResult := E_Result.Passed;
        FExpectedNotInTimespanResult := E_Result.Failed;
        FExpectedFindings := 1;
    LastValidValue:
        FActual := LastValid;
        FReference := LastValid;
        FStart := Zero;
        FEnd := LastValid;
        FExpectedEqualResult := E_Result.Passed;
        FExpectedInTimespanResult := E_Result.Passed;
        FExpectedNotInTimespanResult := E_Result.Failed;
        FExpectedFindings := 1;
    DistinctValid:
        FActual := Zero;
        FReference := LastValid;
        FStart := Zero;
        FEnd := LastValid;
        FExpectedEqualResult := E_Result.Failed;
        FExpectedInTimespanResult := E_Result.Passed;
        FExpectedNotInTimespanResult := E_Result.Failed;
        FExpectedFindings := 2;
    InvalidInput:
        FActual := OneDay;
        FReference := Zero;
        FStart := Zero;
        FEnd := LastValid;
        FExpectedEqualResult := E_Result.Error;
        FExpectedInTimespanResult := E_Result.Error;
        FExpectedNotInTimespanResult := E_Result.Error;
        FExpectedFindings := 3;
    InvalidExpected:
        FActual := Zero;
        FReference := OneDay;
        FStart := Zero;
        FEnd := LastValid;
        FExpectedEqualResult := E_Result.Error;
        FExpectedInTimespanResult := E_Result.Passed;
        FExpectedNotInTimespanResult := E_Result.Failed;
        FExpectedFindings := 2;
    InvalidStart:
        FActual := Zero;
        FReference := Zero;
        FStart := OneDay;
        FEnd := LastValid;
        FExpectedEqualResult := E_Result.Passed;
        FExpectedInTimespanResult := E_Result.Error;
        FExpectedNotInTimespanResult := E_Result.Error;
        FExpectedFindings := 2;
    InvalidEnd:
        FActual := Zero;
        FReference := Zero;
        FStart := Zero;
        FEnd := OneDay;
        FExpectedEqualResult := E_Result.Passed;
        FExpectedInTimespanResult := E_Result.Error;
        FExpectedNotInTimespanResult := E_Result.Error;
        FExpectedFindings := 2;
    ReversedValidSpan:
        FActual := Zero;
        FReference := Zero;
        FStart := LastValid;
        FEnd := Zero;
        FExpectedEqualResult := E_Result.Passed;
        FExpectedInTimespanResult := E_Result.Error;
        FExpectedNotInTimespanResult := E_Result.Error;
        FExpectedFindings := 2;
ELSE
    Error(Message := 'Unknown comparison test row.');
END_CASE;
END_METHOD

END_FUNCTION_BLOCK

// ---- SelfTests/TestCases/TestSuite_AssertionComparisons/Test_AssertionLTODDomain.TcPOU
{region 'Documentation'}
(*!
<summary>Checks all LTOD inputs at midnight and the exclusive 24-hour domain limit.</summary>
<description>
Named rows separate independent comparisons by a disabled reset call.
Only explicitly marked escalation rows retain the preceding subject result.
Outer Assertions latch every observation before advancing to the next row.
Intentional findings remain in the local capture; no production algorithm is copied.
</description>
*)
{endregion}
FUNCTION_BLOCK Test_AssertionLTODDomain EXTENDS TestCaseBase
VAR
    FEqualSubject : AssertEqual_LTOD;
    FInTimespanSubject : AssertInTimespan_LTOD;
    FNotInTimespanSubject : AssertNotInTimespan_LTOD;
    FActual : LTOD;
    FReference : LTOD;
    FStart : LTOD;
    FEnd : LTOD;
    FExpectedEqualResult : E_Result;
    FExpectedInTimespanResult : E_Result;
    FExpectedNotInTimespanResult : E_Result;
    FExpectedFindings : UDINT;
    FCapture : EventBuffer;
    FEvents : ARRAY[1..CaptureLength] OF ST_Event;
    FCaptureFifo : ST_FifoStatus;
    FCaptureStatus : ST_EventBufferStatus;
    FRow : UINT;
    FRowPrepared : BOOL;
    FPreserveResults : BOOL;
    FObservationReady : BOOL;
    FChecked : BOOL;
    FSetupValid : BOOL;
END_VAR
VAR
    FEqualResult : AssertTrue;
    FEqualResultMatches : BOOL;
    FInTimespanResult : AssertTrue;
    FInTimespanResultMatches : BOOL;
    FNotInTimespanResult : AssertTrue;
    FNotInTimespanResultMatches : BOOL;
    FCaptureIntegrity : AssertTrue;
    FCaptureIntegrityMatches : BOOL;
END_VAR
VAR CONSTANT
    CaptureLength : UINT := 8;
    Midnight : UINT := 1;
    LastValidValue : UINT := 2;
    DistinctValid : UINT := 3;
    InvalidInput : UINT := 4;
    InvalidExpected : UINT := 5;
    InvalidStart : UINT := 6;
    InvalidEnd : UINT := 7;
    ReversedValidSpan : UINT := 8;
    LastRow : UINT := ReversedValidSpan;
    Zero : LTOD := LTOD#00:00:00;
    LastValid : LTOD := LTOD#23:59:59.999999999;
    OneDay : LTOD := ULINT_TO_LTOD(ULINT#86400000000000);
END_VAR

SUPER^();

{region 'Documentation'}
(*!
<summary>Collects only outer checking Assertions, never intentional subject findings.</summary>
*)
{endregion}
METHOD PROTECTED AggregateResults
VAR_INPUT
    Aggregator : I_ResultAggregator; //! Borrowed result sink owned by the outer Test Case; add this test's checking Assertions without resetting or retaining the sink.
END_VAR
Aggregator.AddProvider(Provider := FEqualResult);
Aggregator.AddProvider(Provider := FInTimespanResult);
Aggregator.AddProvider(Provider := FNotInTimespanResult);
Aggregator.AddProvider(Provider := FCaptureIntegrity);
END_METHOD

{region 'Documentation'}
(*!
<summary>Calls each inherited production Assertion once using the selected row.</summary>
*)
{endregion}
METHOD PRIVATE CallSubjects
VAR_INPUT
    Enable : BOOL; //! Observation-enable input forwarded to the controlled Assertion subjects for this call.
END_VAR
FEqualSubject(Enable := Enable,
    State := E_State.Running,
    IN := FActual,
    Expected := FReference);
FInTimespanSubject(Enable := Enable,
    State := E_State.Running,
    IN := FActual,
    StartTime := FStart,
    EndTime := FEnd);
FNotInTimespanSubject(Enable := Enable,
    State := E_State.Running,
    IN := FActual,
    StartTime := FStart,
    EndTime := FEnd);
END_METHOD

{region 'Documentation'}
(*!
<summary>Extends base validation with subject and checking-Assertion setup.</summary>
*)
{endregion}
METHOD PROTECTED CheckInitialization : BOOL //! TRUE when the inherited initialization check and this concrete fixture check both accept the setup.
CheckInitialization := SUPER^.CheckInitialization();
IF NOT CheckInitialization THEN
    RETURN;
END_IF;

CheckInitialization := FSetupValid
    AND FEqualResult.IsInitialized
    AND FInTimespanResult.IsInitialized
    AND FNotInTimespanResult.IsInitialized
    AND FCaptureIntegrity.IsInitialized;
IF NOT CheckInitialization THEN
    EventPublisher.PublishEvent(Event := CreateFrameworkEvent(Name := Name,
        ResourceName := '',
        State := State,
        Severity := E_EventSeverity.Error,
        Message := 'Comparison selftest setup failed.'));
END_IF;
END_METHOD

{region 'Documentation'}
(*!
<summary>Checks results and isolated findings against explicit expectations.</summary>
*)
{endregion}
METHOD PRIVATE CheckResults
FEqualResultMatches := FEqualSubject.Result = FExpectedEqualResult;
FInTimespanResultMatches := FInTimespanSubject.Result = FExpectedInTimespanResult;
FNotInTimespanResultMatches := FNotInTimespanSubject.Result = FExpectedNotInTimespanResult;
FCaptureIntegrityMatches := (FCaptureStatus.SequenceId = FExpectedFindings)
    AND (FCaptureStatus.LostEventCount = 0);
END_METHOD

{region 'Documentation'}
(*!
<summary>Configures checking Assertions; subject actions remain in the test script.</summary>
*)
{endregion}
METHOD PROTECTED Configure
VAR
    Initialized : BOOL;
END_VAR
FPreparationStateCount := 0;
FTestStateCount := 1;
FEqualResult.Initialize(Parent := THIS^,
    AssertionName := 'EqualResult');
FInTimespanResult.Initialize(Parent := THIS^,
    AssertionName := 'InTimespanResult');
FNotInTimespanResult.Initialize(Parent := THIS^,
    AssertionName := 'NotInTimespanResult');
FCaptureIntegrity.Initialize(Parent := THIS^,
    AssertionName := 'CaptureIntegrity');
FSetupValid := FCapture.Initialize(Buffer := FEvents,
    FifoControl := FCaptureFifo,
    Status := FCaptureStatus);
FEqualSubject.BindPublisher(Publisher := FCapture);
Initialized := FEqualSubject.Initialize(Parent := THIS^,
    AssertionName := 'EqualSubject');
FSetupValid := FSetupValid AND Initialized;
FInTimespanSubject.BindPublisher(Publisher := FCapture);
Initialized := FInTimespanSubject.Initialize(Parent := THIS^,
    AssertionName := 'InTimespanSubject');
FSetupValid := FSetupValid AND Initialized;
FNotInTimespanSubject.BindPublisher(Publisher := FCapture);
Initialized := FNotInTimespanSubject.Initialize(Parent := THIS^,
    AssertionName := 'NotInTimespanSubject');
FSetupValid := FSetupValid AND Initialized;
END_METHOD

{region 'Documentation'}
(*!
<summary>Completes abort without asynchronous resources.</summary>
*)
{endregion}
METHOD PROTECTED ProcessAbort
VAR_INPUT
    Enable : BOOL; //! Phase permission supplied by the owning Test Case; FALSE does not authorize progression, while observation may continue.
END_VAR
IF Enable THEN
    CompleteAbort();
END_IF;
END_METHOD

{region 'Documentation'}
(*!
<summary>Latches checked observations before the next script step may proceed.</summary>
*)
{endregion}
METHOD PROTECTED ProcessAssertions
VAR_INPUT
    Enable : BOOL; //! Phase permission supplied by the owning Test Case; FALSE does not authorize progression, while observation may continue.
END_VAR
VAR
    Evaluate : BOOL;
END_VAR
Evaluate := Enable AND FObservationReady;
FEqualResult(Enable := Evaluate,
    State := State,
    IN := FEqualResultMatches);
FInTimespanResult(Enable := Evaluate,
    State := State,
    IN := FInTimespanResultMatches);
FNotInTimespanResult(Enable := Evaluate,
    State := State,
    IN := FNotInTimespanResultMatches);
FCaptureIntegrity(Enable := Evaluate,
    State := State,
    IN := FCaptureIntegrityMatches);
IF Evaluate THEN
    FChecked := TRUE;
END_IF;
END_METHOD

{region 'Documentation'}
(*!
<summary>No Preparation phase is required.</summary>
*)
{endregion}
METHOD PROTECTED ProcessPreparations
VAR_INPUT
    // SA0033: Required hook; this test has no Preparation phase.
    {attribute 'analysis' := '-33'}
    Enable : BOOL; //! Phase permission supplied by the owning Test Case; FALSE does not authorize progression, while observation may continue.
END_VAR
END_METHOD

{region 'Documentation'}
(*!
<summary>Restarts the script and resets the checking Assertions.</summary>
*)
{endregion}
METHOD PROTECTED ProcessReset
FRow := Midnight;
FRowPrepared := FALSE;
FChecked := FALSE;
FObservationReady := FALSE;
FEqualResult.Reset();
FEqualResultMatches := TRUE;
FInTimespanResult.Reset();
FInTimespanResultMatches := TRUE;
FNotInTimespanResult.Reset();
FNotInTimespanResultMatches := TRUE;
FCaptureIntegrity.Reset();
FCaptureIntegrityMatches := TRUE;
CompleteReset();
END_METHOD

{region 'Documentation'}
(*!
<summary>Advances one bounded script step per active PLC cycle.</summary>
*)
{endregion}
METHOD PROTECTED ProcessTests
VAR_INPUT
    Enable : BOOL; //! Phase permission supplied by the owning Test Case; FALSE does not authorize progression, while observation may continue.
END_VAR
IF NOT Enable THEN
    RETURN;
END_IF;

IF FChecked THEN
    FChecked := FALSE;
    FObservationReady := FALSE;
    IF FRow = LastRow THEN
        CompleteTests();
        RETURN;
    END_IF;
    FRow := FRow + 1;
    FRowPrepared := FALSE;
END_IF;

IF NOT FRowPrepared THEN
    SelectRow();
    FCapture.Reset();
    IF NOT FPreserveResults THEN
        ResetSubjects();
    END_IF;
    CallSubjects(Enable := FALSE);
    FRowPrepared := TRUE;
ELSE
    CallSubjects(Enable := TRUE);
    CheckResults();
    FObservationReady := TRUE;
END_IF;
END_METHOD

{region 'Documentation'}
(*!
<summary>Requests fresh subject results before the next disabled call.</summary>
*)
{endregion}
METHOD PRIVATE ResetSubjects
FEqualSubject.Reset();
FInTimespanSubject.Reset();
FNotInTimespanSubject.Reset();
END_METHOD

{region 'Documentation'}
(*!
<summary>Selects literal expectations; only named escalation rows retain preceding subject results.</summary>
*)
{endregion}
METHOD PRIVATE SelectRow
FPreserveResults := FALSE;
CASE FRow OF
    Midnight:
        FActual := Zero;
        FReference := Zero;
        FStart := Zero;
        FEnd := LastValid;
        FExpectedEqualResult := E_Result.Passed;
        FExpectedInTimespanResult := E_Result.Passed;
        FExpectedNotInTimespanResult := E_Result.Failed;
        FExpectedFindings := 1;
    LastValidValue:
        FActual := LastValid;
        FReference := LastValid;
        FStart := Zero;
        FEnd := LastValid;
        FExpectedEqualResult := E_Result.Passed;
        FExpectedInTimespanResult := E_Result.Passed;
        FExpectedNotInTimespanResult := E_Result.Failed;
        FExpectedFindings := 1;
    DistinctValid:
        FActual := Zero;
        FReference := LastValid;
        FStart := Zero;
        FEnd := LastValid;
        FExpectedEqualResult := E_Result.Failed;
        FExpectedInTimespanResult := E_Result.Passed;
        FExpectedNotInTimespanResult := E_Result.Failed;
        FExpectedFindings := 2;
    InvalidInput:
        FActual := OneDay;
        FReference := Zero;
        FStart := Zero;
        FEnd := LastValid;
        FExpectedEqualResult := E_Result.Error;
        FExpectedInTimespanResult := E_Result.Error;
        FExpectedNotInTimespanResult := E_Result.Error;
        FExpectedFindings := 3;
    InvalidExpected:
        FActual := Zero;
        FReference := OneDay;
        FStart := Zero;
        FEnd := LastValid;
        FExpectedEqualResult := E_Result.Error;
        FExpectedInTimespanResult := E_Result.Passed;
        FExpectedNotInTimespanResult := E_Result.Failed;
        FExpectedFindings := 2;
    InvalidStart:
        FActual := Zero;
        FReference := Zero;
        FStart := OneDay;
        FEnd := LastValid;
        FExpectedEqualResult := E_Result.Passed;
        FExpectedInTimespanResult := E_Result.Error;
        FExpectedNotInTimespanResult := E_Result.Error;
        FExpectedFindings := 2;
    InvalidEnd:
        FActual := Zero;
        FReference := Zero;
        FStart := Zero;
        FEnd := OneDay;
        FExpectedEqualResult := E_Result.Passed;
        FExpectedInTimespanResult := E_Result.Error;
        FExpectedNotInTimespanResult := E_Result.Error;
        FExpectedFindings := 2;
    ReversedValidSpan:
        FActual := Zero;
        FReference := Zero;
        FStart := LastValid;
        FEnd := Zero;
        FExpectedEqualResult := E_Result.Passed;
        FExpectedInTimespanResult := E_Result.Error;
        FExpectedNotInTimespanResult := E_Result.Error;
        FExpectedFindings := 2;
ELSE
    Error(Message := 'Unknown comparison test row.');
END_CASE;
END_METHOD

END_FUNCTION_BLOCK

// ---- Framework/Assertions/POU/BasicTypes/LTOD/AssertEqual_LTOD.TcPOU
{region 'Documentation'}
(*!
<summary>Checks equality with the expected LTOD value.</summary>
<description>

A value at or beyond 24 hours reports Error before comparison or baseline capture.

</description>
*)
{endregion}
FUNCTION_BLOCK AssertEqual_LTOD EXTENDS AssertionBase
VAR_INPUT
    IN : LTOD; //! Actual value checked or observed by this Assertion.
    Expected : LTOD; //! Reference value for comparison with IN.
END_VAR

SUPER^();

{region 'Documentation'}
(*!
<summary>Evaluate the typed temporal relation and report higher-priority errors first.</summary>
*)
{endregion}
METHOD PROTECTED Assert
VAR
    Message : STRING(GVL_Constants.MessageLength);
    ExpectedText : STRING(GVL_Constants.AssertionValueLength);
    ActualText : STRING(GVL_Constants.AssertionValueLength);
END_VAR
IF NOT EvaluationActive THEN
    RETURN;
END_IF;

IF Result = E_Result.Error THEN
    RETURN;
END_IF;

IF NOT IsTimeOfDayValid_LTOD(Value := IN) THEN
    Error(Message := 'Assertion error: IN is outside the valid LTOD range (less than 24 hours).');
    RETURN;
END_IF;

IF NOT IsTimeOfDayValid_LTOD(Value := Expected) THEN
    Error(Message := 'Assertion error: Expected is outside the valid LTOD range (less than 24 hours).');
    RETURN;
END_IF;

IF Result = E_Result.Failed THEN
    RETURN;
END_IF;

IF IN <> Expected THEN
    ExpectedText := LTOD_TO_STRING(Expected);
    ActualText := LTOD_TO_STRING(IN);
    Message := CONCAT('Assertion failed: values are not equal. Expected = ',
        ExpectedText);
    Message := CONCAT(Message, ', Actual = ');
    Message := CONCAT(Message, ActualText);
    Message := CONCAT(Message, '.');
    Fail(Message := Message);
    RETURN;
END_IF;

Pass();
END_METHOD

END_FUNCTION_BLOCK

// ---- Framework/Assertions/POU/Utilities/IsTimeOfDayValid_LTOD.TcPOU
{region 'Documentation'}
(*!
<summary>Checks the native time-of-day range without changing or normalizing Value.</summary>
*)
{endregion}
FUNCTION INTERNAL IsTimeOfDayValid_LTOD : BOOL //! TRUE for a time of day below 24 hours; the value is not normalized.
VAR_INPUT
    Value : LTOD; //! Time-of-day value checked against the interval from midnight inclusive to the next midnight exclusive.
END_VAR
VAR CONSTANT
    MaximumTimeOfDay : LTOD := LTOD#23:59:59.999999999;
END_VAR

IsTimeOfDayValid_LTOD := Value <= MaximumTimeOfDay;

END_FUNCTION

// ---- Framework/Assertions/POU/BasicTypes/LTOD/AssertInTimespan_LTOD.TcPOU
{region 'Documentation'}
(*!
<summary>Check that IN is inside the inclusive StartTime..EndTime interval.</summary>
<description>

StartTime &gt; EndTime reports Error during active evaluation; equal bounds are
valid.

A value at or beyond 24 hours reports Error before comparison or baseline capture.

</description>
*)
{endregion}
FUNCTION_BLOCK AssertInTimespan_LTOD EXTENDS AssertionBase
VAR_INPUT
    IN : LTOD; //! Actual value checked or observed by this Assertion.
    StartTime : LTOD; //! Inclusive start of the time span; must not exceed EndTime.
    EndTime : LTOD; //! Inclusive end of the time span; must not precede StartTime.
END_VAR

SUPER^();

{region 'Documentation'}
(*!
<summary>Evaluate the typed temporal relation and report higher-priority errors first.</summary>
*)
{endregion}
METHOD PROTECTED Assert
VAR
    Message : STRING(GVL_Constants.MessageLength);
    StartTimeText : STRING(GVL_Constants.AssertionValueLength);
    EndTimeText : STRING(GVL_Constants.AssertionValueLength);
    ActualText : STRING(GVL_Constants.AssertionValueLength);
END_VAR
IF NOT EvaluationActive THEN
    RETURN;
END_IF;

IF Result = E_Result.Error THEN
    RETURN;
END_IF;

IF NOT IsTimeOfDayValid_LTOD(Value := IN) THEN
    Error(Message := 'Assertion error: IN is outside the valid LTOD range (less than 24 hours).');
    RETURN;
END_IF;

IF NOT IsTimeOfDayValid_LTOD(Value := StartTime) THEN
    Error(Message := 'Assertion error: StartTime is outside the valid LTOD range (less than 24 hours).');
    RETURN;
END_IF;

IF NOT IsTimeOfDayValid_LTOD(Value := EndTime) THEN
    Error(Message := 'Assertion error: EndTime is outside the valid LTOD range (less than 24 hours).');
    RETURN;
END_IF;

IF StartTime > EndTime THEN
    StartTimeText := LTOD_TO_STRING(StartTime);
    EndTimeText := LTOD_TO_STRING(EndTime);
    Message := CONCAT('Assertion error: start time exceeds end time. StartTime = ',
        StartTimeText);
    Message := CONCAT(Message, ', EndTime = ');
    Message := CONCAT(Message, EndTimeText);
    Message := CONCAT(Message, '.');
    Error(Message := Message);
    RETURN;
END_IF;

IF Result = E_Result.Failed THEN
    RETURN;
END_IF;

IF (IN < StartTime) OR (IN > EndTime) THEN
    StartTimeText := LTOD_TO_STRING(StartTime);
    EndTimeText := LTOD_TO_STRING(EndTime);
    ActualText := LTOD_TO_STRING(IN);
    Message := CONCAT('Assertion failed: value is outside allowed timespan. StartTime = ',
        StartTimeText);
    Message := CONCAT(Message, ', EndTime = ');
    Message := CONCAT(Message, EndTimeText);
    Message := CONCAT(Message, ', Actual = ');
    Message := CONCAT(Message, ActualText);
    Message := CONCAT(Message, '.');
    Fail(Message := Message);
    RETURN;
END_IF;

Pass();
END_METHOD

END_FUNCTION_BLOCK

// ---- Framework/Assertions/POU/BasicTypes/LTOD/AssertNotInTimespan_LTOD.TcPOU
{region 'Documentation'}
(*!
<summary>Check that IN is outside the inclusive StartTime..EndTime interval.</summary>
<description>

StartTime &gt; EndTime reports Error during active evaluation; equal bounds are
valid.

A value at or beyond 24 hours reports Error before comparison or baseline capture.

</description>
*)
{endregion}
FUNCTION_BLOCK AssertNotInTimespan_LTOD EXTENDS AssertionBase
VAR_INPUT
    IN : LTOD; //! Actual value checked or observed by this Assertion.
    StartTime : LTOD; //! Inclusive start of the time span; must not exceed EndTime.
    EndTime : LTOD; //! Inclusive end of the time span; must not precede StartTime.
END_VAR

SUPER^();

{region 'Documentation'}
(*!
<summary>Evaluate the typed temporal relation and report higher-priority errors first.</summary>
*)
{endregion}
METHOD PROTECTED Assert
VAR
    Message : STRING(GVL_Constants.MessageLength);
    StartTimeText : STRING(GVL_Constants.AssertionValueLength);
    EndTimeText : STRING(GVL_Constants.AssertionValueLength);
    ActualText : STRING(GVL_Constants.AssertionValueLength);
END_VAR
IF NOT EvaluationActive THEN
    RETURN;
END_IF;

IF Result = E_Result.Error THEN
    RETURN;
END_IF;

IF NOT IsTimeOfDayValid_LTOD(Value := IN) THEN
    Error(Message := 'Assertion error: IN is outside the valid LTOD range (less than 24 hours).');
    RETURN;
END_IF;

IF NOT IsTimeOfDayValid_LTOD(Value := StartTime) THEN
    Error(Message := 'Assertion error: StartTime is outside the valid LTOD range (less than 24 hours).');
    RETURN;
END_IF;

IF NOT IsTimeOfDayValid_LTOD(Value := EndTime) THEN
    Error(Message := 'Assertion error: EndTime is outside the valid LTOD range (less than 24 hours).');
    RETURN;
END_IF;

IF StartTime > EndTime THEN
    StartTimeText := LTOD_TO_STRING(StartTime);
    EndTimeText := LTOD_TO_STRING(EndTime);
    Message := CONCAT('Assertion error: start time exceeds end time. StartTime = ',
        StartTimeText);
    Message := CONCAT(Message, ', EndTime = ');
    Message := CONCAT(Message, EndTimeText);
    Message := CONCAT(Message, '.');
    Error(Message := Message);
    RETURN;
END_IF;

IF Result = E_Result.Failed THEN
    RETURN;
END_IF;

IF (IN >= StartTime) AND (IN <= EndTime) THEN
    StartTimeText := LTOD_TO_STRING(StartTime);
    EndTimeText := LTOD_TO_STRING(EndTime);
    ActualText := LTOD_TO_STRING(IN);
    Message := CONCAT('Assertion failed: value is inside forbidden timespan. StartTime = ',
        StartTimeText);
    Message := CONCAT(Message, ', EndTime = ');
    Message := CONCAT(Message, EndTimeText);
    Message := CONCAT(Message, ', Actual = ');
    Message := CONCAT(Message, ActualText);
    Message := CONCAT(Message, '.');
    Fail(Message := Message);
    RETURN;
END_IF;

Pass();
END_METHOD

END_FUNCTION_BLOCK

// ---- SelfTests/TestCases/TestSuite_AssertionComparisons/Test_AssertionScalarDiagnostics.TcPOU
{region 'Documentation'}
(*!
<summary>Checks literal expected/actual decimal, fixed-width hex and character rendering in captured findings.</summary>
<description>
Named rows separate independent comparisons by a disabled reset call.
Only explicitly marked escalation rows retain the preceding subject result.
Outer Assertions latch every observation before advancing to the next row.
Intentional findings remain in the local capture; no production algorithm is copied.
</description>
*)
{endregion}
FUNCTION_BLOCK Test_AssertionScalarDiagnostics EXTENDS TestCaseBase
VAR
    FSignedSubject : AssertEqual_LInt;
    FUnsignedSubject : AssertEqual_ULInt;
    FByteSubject : AssertEqual_Byte;
    FLWordSubject : AssertEqual_LWord;
    FCharSubject : AssertEqual_Char;
    FWCharSubject : AssertEqual_WChar;
    FActualSigned : LINT;
    FReferenceSigned : LINT;
    FExpectedSignedMessage : STRING(GVL_Constants.MessageLength);
    FActualUnsigned : ULINT;
    FReferenceUnsigned : ULINT;
    FExpectedUnsignedMessage : STRING(GVL_Constants.MessageLength);
    FActualByte : BYTE;
    FReferenceByte : BYTE;
    FExpectedByteMessage : STRING(GVL_Constants.MessageLength);
    FActualLWord : LWORD;
    FReferenceLWord : LWORD;
    FExpectedLWordMessage : STRING(GVL_Constants.MessageLength);
    FActualChar : BYTE;
    FReferenceChar : BYTE;
    FExpectedCharMessage : STRING(GVL_Constants.MessageLength);
    FActualWChar : WORD;
    FReferenceWChar : WORD;
    FExpectedWCharMessage : STRING(GVL_Constants.MessageLength);
    FExpectedSignedResult : E_Result;
    FExpectedUnsignedResult : E_Result;
    FExpectedByteResult : E_Result;
    FExpectedLWordResult : E_Result;
    FExpectedCharResult : E_Result;
    FExpectedWCharResult : E_Result;
    FExpectedFindings : UDINT;
    FCapture : EventBuffer;
    FEvents : ARRAY[1..CaptureLength] OF ST_Event;
    FCaptureFifo : ST_FifoStatus;
    FCaptureStatus : ST_EventBufferStatus;
    FRow : UINT;
    FRowPrepared : BOOL;
    FPreserveResults : BOOL;
    FObservationReady : BOOL;
    FChecked : BOOL;
    FSetupValid : BOOL;
END_VAR
VAR
    FSignedResult : AssertTrue;
    FSignedResultMatches : BOOL;
    FUnsignedResult : AssertTrue;
    FUnsignedResultMatches : BOOL;
    FByteResult : AssertTrue;
    FByteResultMatches : BOOL;
    FLWordResult : AssertTrue;
    FLWordResultMatches : BOOL;
    FCharResult : AssertTrue;
    FCharResultMatches : BOOL;
    FWCharResult : AssertTrue;
    FWCharResultMatches : BOOL;
    FCaptureIntegrity : AssertTrue;
    FCaptureIntegrityMatches : BOOL;
    FDiagnosticText : AssertTrue;
    FDiagnosticTextMatches : BOOL;
END_VAR
VAR CONSTANT
    CaptureLength : UINT := 16;
    Printable : UINT := 1;
    NullAndWide : UINT := 2;
    MaximumCodes : UINT := 3;
    LastRow : UINT := MaximumCodes;

END_VAR

SUPER^();

{region 'Documentation'}
(*!
<summary>Collects only outer checking Assertions, never intentional subject findings.</summary>
*)
{endregion}
METHOD PROTECTED AggregateResults
VAR_INPUT
    Aggregator : I_ResultAggregator; //! Borrowed result sink owned by the outer Test Case; add this test's checking Assertions without resetting or retaining the sink.
END_VAR
Aggregator.AddProvider(Provider := FSignedResult);
Aggregator.AddProvider(Provider := FUnsignedResult);
Aggregator.AddProvider(Provider := FByteResult);
Aggregator.AddProvider(Provider := FLWordResult);
Aggregator.AddProvider(Provider := FCharResult);
Aggregator.AddProvider(Provider := FWCharResult);
Aggregator.AddProvider(Provider := FCaptureIntegrity);
Aggregator.AddProvider(Provider := FDiagnosticText);
END_METHOD

{region 'Documentation'}
(*!
<summary>Calls each inherited production Assertion once using the selected row.</summary>
*)
{endregion}
METHOD PRIVATE CallSubjects
VAR_INPUT
    Enable : BOOL; //! Observation-enable input forwarded to the controlled Assertion subjects for this call.
END_VAR
FSignedSubject(Enable := Enable,
    State := E_State.Running,
    IN := FActualSigned,
    Expected := FReferenceSigned);
FUnsignedSubject(Enable := Enable,
    State := E_State.Running,
    IN := FActualUnsigned,
    Expected := FReferenceUnsigned);
FByteSubject(Enable := Enable,
    State := E_State.Running,
    IN := FActualByte,
    Expected := FReferenceByte);
FLWordSubject(Enable := Enable,
    State := E_State.Running,
    IN := FActualLWord,
    Expected := FReferenceLWord);
FCharSubject(Enable := Enable,
    State := E_State.Running,
    IN := FActualChar,
    Expected := FReferenceChar);
FWCharSubject(Enable := Enable,
    State := E_State.Running,
    IN := FActualWChar,
    Expected := FReferenceWChar);
END_METHOD

{region 'Documentation'}
(*!
<summary>Extends base validation with subject and checking-Assertion setup.</summary>
*)
{endregion}
METHOD PROTECTED CheckInitialization : BOOL //! TRUE when the inherited initialization check and this concrete fixture check both accept the setup.
CheckInitialization := SUPER^.CheckInitialization();
IF NOT CheckInitialization THEN
    RETURN;
END_IF;

CheckInitialization := FSetupValid
    AND FSignedResult.IsInitialized
    AND FUnsignedResult.IsInitialized
    AND FByteResult.IsInitialized
    AND FLWordResult.IsInitialized
    AND FCharResult.IsInitialized
    AND FWCharResult.IsInitialized
    AND FCaptureIntegrity.IsInitialized
    AND FDiagnosticText.IsInitialized;
IF NOT CheckInitialization THEN
    EventPublisher.PublishEvent(Event := CreateFrameworkEvent(Name := Name,
        ResourceName := '',
        State := State,
        Severity := E_EventSeverity.Error,
        Message := 'Comparison selftest setup failed.'));
END_IF;
END_METHOD

{region 'Documentation'}
(*!
<summary>Checks results and isolated findings against explicit expectations.</summary>
*)
{endregion}
METHOD PRIVATE CheckResults
FSignedResultMatches := FSignedSubject.Result = FExpectedSignedResult;
FUnsignedResultMatches := FUnsignedSubject.Result = FExpectedUnsignedResult;
FByteResultMatches := FByteSubject.Result = FExpectedByteResult;
FLWordResultMatches := FLWordSubject.Result = FExpectedLWordResult;
FCharResultMatches := FCharSubject.Result = FExpectedCharResult;
FWCharResultMatches := FWCharSubject.Result = FExpectedWCharResult;
FCaptureIntegrityMatches := (FCaptureStatus.SequenceId = FExpectedFindings)
    AND (FCaptureStatus.LostEventCount = 0);
FDiagnosticTextMatches := (FEvents[1].Message = FExpectedSignedMessage)
    AND (FEvents[1].Name = FSignedSubject.Name)
    AND (FEvents[1].Result = E_Result.Failed)
    AND (FEvents[2].Message = FExpectedUnsignedMessage)
    AND (FEvents[2].Name = FUnsignedSubject.Name)
    AND (FEvents[2].Result = E_Result.Failed)
    AND (FEvents[3].Message = FExpectedByteMessage)
    AND (FEvents[3].Name = FByteSubject.Name)
    AND (FEvents[3].Result = E_Result.Failed)
    AND (FEvents[4].Message = FExpectedLWordMessage)
    AND (FEvents[4].Name = FLWordSubject.Name)
    AND (FEvents[4].Result = E_Result.Failed)
    AND (FEvents[5].Message = FExpectedCharMessage)
    AND (FEvents[5].Name = FCharSubject.Name)
    AND (FEvents[5].Result = E_Result.Failed)
    AND (FEvents[6].Message = FExpectedWCharMessage)
    AND (FEvents[6].Name = FWCharSubject.Name)
    AND (FEvents[6].Result = E_Result.Failed);
END_METHOD

{region 'Documentation'}
(*!
<summary>Configures checking Assertions; subject actions remain in the test script.</summary>
*)
{endregion}
METHOD PROTECTED Configure
VAR
    Initialized : BOOL;
END_VAR
FPreparationStateCount := 0;
FTestStateCount := 1;
FSignedResult.Initialize(Parent := THIS^,
    AssertionName := 'SignedResult');
FUnsignedResult.Initialize(Parent := THIS^,
    AssertionName := 'UnsignedResult');
FByteResult.Initialize(Parent := THIS^,
    AssertionName := 'ByteResult');
FLWordResult.Initialize(Parent := THIS^,
    AssertionName := 'LWordResult');
FCharResult.Initialize(Parent := THIS^,
    AssertionName := 'CharResult');
FWCharResult.Initialize(Parent := THIS^,
    AssertionName := 'WCharResult');
FCaptureIntegrity.Initialize(Parent := THIS^,
    AssertionName := 'CaptureIntegrity');
FDiagnosticText.Initialize(Parent := THIS^,
    AssertionName := 'DiagnosticText');
FSetupValid := FCapture.Initialize(Buffer := FEvents,
    FifoControl := FCaptureFifo,
    Status := FCaptureStatus);
FSignedSubject.BindPublisher(Publisher := FCapture);
Initialized := FSignedSubject.Initialize(Parent := THIS^,
    AssertionName := 'SignedSubject');
FSetupValid := FSetupValid AND Initialized;
FUnsignedSubject.BindPublisher(Publisher := FCapture);
Initialized := FUnsignedSubject.Initialize(Parent := THIS^,
    AssertionName := 'UnsignedSubject');
FSetupValid := FSetupValid AND Initialized;
FByteSubject.BindPublisher(Publisher := FCapture);
Initialized := FByteSubject.Initialize(Parent := THIS^,
    AssertionName := 'ByteSubject');
FSetupValid := FSetupValid AND Initialized;
FLWordSubject.BindPublisher(Publisher := FCapture);
Initialized := FLWordSubject.Initialize(Parent := THIS^,
    AssertionName := 'LWordSubject');
FSetupValid := FSetupValid AND Initialized;
FCharSubject.BindPublisher(Publisher := FCapture);
Initialized := FCharSubject.Initialize(Parent := THIS^,
    AssertionName := 'CharSubject');
FSetupValid := FSetupValid AND Initialized;
FWCharSubject.BindPublisher(Publisher := FCapture);
Initialized := FWCharSubject.Initialize(Parent := THIS^,
    AssertionName := 'WCharSubject');
FSetupValid := FSetupValid AND Initialized;
END_METHOD

{region 'Documentation'}
(*!
<summary>Completes abort without asynchronous resources.</summary>
*)
{endregion}
METHOD PROTECTED ProcessAbort
VAR_INPUT
    Enable : BOOL; //! Phase permission supplied by the owning Test Case; FALSE does not authorize progression, while observation may continue.
END_VAR
IF Enable THEN
    CompleteAbort();
END_IF;
END_METHOD

{region 'Documentation'}
(*!
<summary>Latches checked observations before the next script step may proceed.</summary>
*)
{endregion}
METHOD PROTECTED ProcessAssertions
VAR_INPUT
    Enable : BOOL; //! Phase permission supplied by the owning Test Case; FALSE does not authorize progression, while observation may continue.
END_VAR
VAR
    Evaluate : BOOL;
END_VAR
Evaluate := Enable AND FObservationReady;
FSignedResult(Enable := Evaluate,
    State := State,
    IN := FSignedResultMatches);
FUnsignedResult(Enable := Evaluate,
    State := State,
    IN := FUnsignedResultMatches);
FByteResult(Enable := Evaluate,
    State := State,
    IN := FByteResultMatches);
FLWordResult(Enable := Evaluate,
    State := State,
    IN := FLWordResultMatches);
FCharResult(Enable := Evaluate,
    State := State,
    IN := FCharResultMatches);
FWCharResult(Enable := Evaluate,
    State := State,
    IN := FWCharResultMatches);
FCaptureIntegrity(Enable := Evaluate,
    State := State,
    IN := FCaptureIntegrityMatches);
FDiagnosticText(Enable := Evaluate,
    State := State,
    IN := FDiagnosticTextMatches);
IF Evaluate THEN
    FChecked := TRUE;
END_IF;
END_METHOD

{region 'Documentation'}
(*!
<summary>No Preparation phase is required.</summary>
*)
{endregion}
METHOD PROTECTED ProcessPreparations
VAR_INPUT
    // SA0033: Required hook; this test has no Preparation phase.
    {attribute 'analysis' := '-33'}
    Enable : BOOL; //! Phase permission supplied by the owning Test Case; FALSE does not authorize progression, while observation may continue.
END_VAR
END_METHOD

{region 'Documentation'}
(*!
<summary>Restarts the script and resets the checking Assertions.</summary>
*)
{endregion}
METHOD PROTECTED ProcessReset
FRow := Printable;
FRowPrepared := FALSE;
FChecked := FALSE;
FObservationReady := FALSE;
FSignedResult.Reset();
FSignedResultMatches := TRUE;
FUnsignedResult.Reset();
FUnsignedResultMatches := TRUE;
FByteResult.Reset();
FByteResultMatches := TRUE;
FLWordResult.Reset();
FLWordResultMatches := TRUE;
FCharResult.Reset();
FCharResultMatches := TRUE;
FWCharResult.Reset();
FWCharResultMatches := TRUE;
FCaptureIntegrity.Reset();
FCaptureIntegrityMatches := TRUE;
FDiagnosticText.Reset();
FDiagnosticTextMatches := TRUE;
CompleteReset();
END_METHOD

{region 'Documentation'}
(*!
<summary>Advances one bounded script step per active PLC cycle.</summary>
*)
{endregion}
METHOD PROTECTED ProcessTests
VAR_INPUT
    Enable : BOOL; //! Phase permission supplied by the owning Test Case; FALSE does not authorize progression, while observation may continue.
END_VAR
IF NOT Enable THEN
    RETURN;
END_IF;

IF FChecked THEN
    FChecked := FALSE;
    FObservationReady := FALSE;
    IF FRow = LastRow THEN
        CompleteTests();
        RETURN;
    END_IF;
    FRow := FRow + 1;
    FRowPrepared := FALSE;
END_IF;

IF NOT FRowPrepared THEN
    SelectRow();
    FCapture.Reset();
    IF NOT FPreserveResults THEN
        ResetSubjects();
    END_IF;
    CallSubjects(Enable := FALSE);
    FRowPrepared := TRUE;
ELSE
    CallSubjects(Enable := TRUE);
    CheckResults();
    FObservationReady := TRUE;
END_IF;
END_METHOD

{region 'Documentation'}
(*!
<summary>Requests fresh subject results before the next disabled call.</summary>
*)
{endregion}
METHOD PRIVATE ResetSubjects
FSignedSubject.Reset();
FUnsignedSubject.Reset();
FByteSubject.Reset();
FLWordSubject.Reset();
FCharSubject.Reset();
FWCharSubject.Reset();
END_METHOD

{region 'Documentation'}
(*!
<summary>Selects literal expectations; only named escalation rows retain preceding subject results.</summary>
*)
{endregion}
METHOD PRIVATE SelectRow
FPreserveResults := FALSE;
CASE FRow OF
    Printable:
        FActualSigned := LINT#-9223372036854775808;
        FReferenceSigned := LINT#9223372036854775807;
        FActualUnsigned := ULINT#18446744073709551615;
        FReferenceUnsigned := ULINT#0;
        FActualByte := BYTE#16#80;
        FReferenceByte := BYTE#16#01;
        FActualLWord := LWORD#16#8000000000000000;
        FReferenceLWord := LWORD#16#0000000000000001;
        FActualChar := BYTE#16#41;
        FReferenceChar := BYTE#16#42;
        FActualWChar := WORD#16#0041;
        FReferenceWChar := WORD#16#0042;
        FExpectedSignedMessage := 'Assertion failed: values are not equal. Expected = 9223372036854775807, Actual = -9223372036854775808.';
        FExpectedUnsignedMessage := 'Assertion failed: values are not equal. Expected = 0, Actual = 18446744073709551615.';
        FExpectedByteMessage := 'Assertion failed: values are not equal. Expected = 16#01, Actual = 16#80.';
        FExpectedLWordMessage := 'Assertion failed: values are not equal. Expected = 16#0000000000000001, Actual = 16#8000000000000000.';
        FExpectedCharMessage := 'Assertion failed: values are not equal. Expected = $'B$' (16#42), Actual = $'A$' (16#41).';
        FExpectedWCharMessage := 'Assertion failed: values are not equal. Expected = $'B$' (16#0042), Actual = $'A$' (16#0041).';
        FExpectedSignedResult := E_Result.Failed;
        FExpectedUnsignedResult := E_Result.Failed;
        FExpectedByteResult := E_Result.Failed;
        FExpectedLWordResult := E_Result.Failed;
        FExpectedCharResult := E_Result.Failed;
        FExpectedWCharResult := E_Result.Failed;
        FExpectedFindings := 6;
    NullAndWide:
        FActualSigned := LINT#-9223372036854775808;
        FReferenceSigned := LINT#9223372036854775807;
        FActualUnsigned := ULINT#18446744073709551615;
        FReferenceUnsigned := ULINT#0;
        FActualByte := BYTE#16#80;
        FReferenceByte := BYTE#16#01;
        FActualLWord := LWORD#16#8000000000000000;
        FReferenceLWord := LWORD#16#0000000000000001;
        FActualChar := BYTE#0;
        FReferenceChar := BYTE#16#41;
        FActualWChar := WORD#16#0100;
        FReferenceWChar := WORD#0;
        FExpectedSignedMessage := 'Assertion failed: values are not equal. Expected = 9223372036854775807, Actual = -9223372036854775808.';
        FExpectedUnsignedMessage := 'Assertion failed: values are not equal. Expected = 0, Actual = 18446744073709551615.';
        FExpectedByteMessage := 'Assertion failed: values are not equal. Expected = 16#01, Actual = 16#80.';
        FExpectedLWordMessage := 'Assertion failed: values are not equal. Expected = 16#0000000000000001, Actual = 16#8000000000000000.';
        FExpectedCharMessage := 'Assertion failed: values are not equal. Expected = $'A$' (16#41), Actual = 16#00.';
        FExpectedWCharMessage := 'Assertion failed: values are not equal. Expected = 16#0000, Actual = 16#0100.';
        FExpectedSignedResult := E_Result.Failed;
        FExpectedUnsignedResult := E_Result.Failed;
        FExpectedByteResult := E_Result.Failed;
        FExpectedLWordResult := E_Result.Failed;
        FExpectedCharResult := E_Result.Failed;
        FExpectedWCharResult := E_Result.Failed;
        FExpectedFindings := 6;
    MaximumCodes:
        FActualSigned := LINT#-9223372036854775808;
        FReferenceSigned := LINT#9223372036854775807;
        FActualUnsigned := ULINT#18446744073709551615;
        FReferenceUnsigned := ULINT#0;
        FActualByte := BYTE#16#80;
        FReferenceByte := BYTE#16#01;
        FActualLWord := LWORD#16#8000000000000000;
        FReferenceLWord := LWORD#16#0000000000000001;
        FActualChar := BYTE#16#FF;
        FReferenceChar := BYTE#0;
        FActualWChar := WORD#16#FFFF;
        FReferenceWChar := WORD#0;
        FExpectedSignedMessage := 'Assertion failed: values are not equal. Expected = 9223372036854775807, Actual = -9223372036854775808.';
        FExpectedUnsignedMessage := 'Assertion failed: values are not equal. Expected = 0, Actual = 18446744073709551615.';
        FExpectedByteMessage := 'Assertion failed: values are not equal. Expected = 16#01, Actual = 16#80.';
        FExpectedLWordMessage := 'Assertion failed: values are not equal. Expected = 16#0000000000000001, Actual = 16#8000000000000000.';
        FExpectedCharMessage := 'Assertion failed: values are not equal. Expected = 16#00, Actual = 16#FF.';
        FExpectedWCharMessage := 'Assertion failed: values are not equal. Expected = 16#0000, Actual = 16#FFFF.';
        FExpectedSignedResult := E_Result.Failed;
        FExpectedUnsignedResult := E_Result.Failed;
        FExpectedByteResult := E_Result.Failed;
        FExpectedLWordResult := E_Result.Failed;
        FExpectedCharResult := E_Result.Failed;
        FExpectedWCharResult := E_Result.Failed;
        FExpectedFindings := 6;
ELSE
    Error(Message := 'Unknown comparison test row.');
END_CASE;
END_METHOD

END_FUNCTION_BLOCK

// ---- SelfTests/TestSuites/TestSuite_AssertionFloatingPoint.TcPOU
{region 'Documentation'}
(*!
<summary>Checks floating-point tolerances, finite boundaries, scalar/array classification and non-finite diagnostics.</summary>
*)
{endregion}
FUNCTION_BLOCK TestSuite_AssertionFloatingPoint EXTENDS TestSuiteBase
VAR
    FTolerance_Real : Test_AssertionTolerance_Real;
    FTolerance_LReal : Test_AssertionTolerance_LReal;
    FFiniteBoundaries_Real : Test_AssertionFiniteBoundaries_Real;
    FFiniteBoundaries_LReal : Test_AssertionFiniteBoundaries_LReal;
    FRelations_Real : Test_AssertionRelations_Real;
    FRelations_LReal : Test_AssertionRelations_LReal;
    FNonFinite_Real : Test_AssertionNonFinite_Real;
    FNonFinite_LReal : Test_AssertionNonFinite_LReal;
    FTestCases : ARRAY[1..TestCaseCapacity] OF I_TestCase;
    FClassification_Real : Test_AssertionClassification_Real;
    FArrayClassification_Real : Test_AssertionArrayClassification_Real;
    FClassification_LReal : Test_AssertionClassification_LReal;
    FArrayClassification_LReal : Test_AssertionArrayClassification_LReal;
END_VAR
VAR CONSTANT
    TestCaseCapacity : UINT := 12;
END_VAR

SUPER^();

{region 'Documentation'}
(*!
<summary>Initializes and registers the twelve isolated floating-point scenarios.</summary>
*)
{endregion}
METHOD PROTECTED Configure
VAR_IN_OUT
    // SA0167: Borrowed owner builder; no temporary instance is created.
    {attribute 'analysis' := '-167'}
    Builder : TestSuiteConfigurationBuilder; //! Borrowed owner configuration builder used only during this Configure call; register this owner's concrete children.
END_VAR
VAR
    TestConfig : ST_TestCaseConfig;
END_VAR
Builder.Initialize(Mode := E_OrchestrationMode.Serial,
    TestCases := FTestCases);
FTolerance_Real.Initialize(Parent := THIS^,
    TestName := 'Tolerance_Real',
    Config := TestConfig);
Builder.Register(TestCase := FTolerance_Real);
FTolerance_LReal.Initialize(Parent := THIS^,
    TestName := 'Tolerance_LReal',
    Config := TestConfig);
Builder.Register(TestCase := FTolerance_LReal);
FFiniteBoundaries_Real.Initialize(Parent := THIS^,
    TestName := 'FiniteBoundaries_Real',
    Config := TestConfig);
Builder.Register(TestCase := FFiniteBoundaries_Real);
FFiniteBoundaries_LReal.Initialize(Parent := THIS^,
    TestName := 'FiniteBoundaries_LReal',
    Config := TestConfig);
Builder.Register(TestCase := FFiniteBoundaries_LReal);
FRelations_Real.Initialize(Parent := THIS^,
    TestName := 'Relations_Real',
    Config := TestConfig);
Builder.Register(TestCase := FRelations_Real);
FRelations_LReal.Initialize(Parent := THIS^,
    TestName := 'Relations_LReal',
    Config := TestConfig);
Builder.Register(TestCase := FRelations_LReal);
FNonFinite_Real.Initialize(Parent := THIS^,
    TestName := 'NonFinite_Real',
    Config := TestConfig);
Builder.Register(TestCase := FNonFinite_Real);
FNonFinite_LReal.Initialize(Parent := THIS^,
    TestName := 'NonFinite_LReal',
    Config := TestConfig);
Builder.Register(TestCase := FNonFinite_LReal);

FClassification_Real.Initialize(Parent := THIS^,
    TestName := 'Classify_Real',
    Config := TestConfig);
Builder.Register(TestCase := FClassification_Real);
FArrayClassification_Real.Initialize(Parent := THIS^,
    TestName := 'ArrayClassify_Real',
    Config := TestConfig);
Builder.Register(TestCase := FArrayClassification_Real);
FClassification_LReal.Initialize(Parent := THIS^,
    TestName := 'Classify_LReal',
    Config := TestConfig);
Builder.Register(TestCase := FClassification_LReal);
FArrayClassification_LReal.Initialize(Parent := THIS^,
    TestName := 'ArrayClassify_LReal',
    Config := TestConfig);
Builder.Register(TestCase := FArrayClassification_LReal);
END_METHOD

{region 'Documentation'}
(*!
<summary>Returns a registered scenario using its original array index.</summary>
*)
{endregion}
METHOD PUBLIC GetTestCase : I_TestCase //! Typed child interface at the original array index; zero when no entry is available.
VAR_INPUT
    Index : DINT; //! Original occupied child-array index, rather than an ordinal position.
END_VAR
GetTestCase := 0;
IF (ChildCount = 0) OR (Index < ChildArrayLowerBound)
    OR (DINT_TO_LINT(Index) >= DINT_TO_LINT(ChildArrayLowerBound) + UINT_TO_LINT(ChildCount)) THEN
    RETURN;
END_IF;
GetTestCase := FTestCases[Index];
END_METHOD

{region 'Documentation'}
(*!
<summary>Calls each owned scenario once per initialized Suite cycle.</summary>
*)
{endregion}
METHOD PROTECTED ProcessTestCases
FTolerance_Real();
FTolerance_LReal();
FFiniteBoundaries_Real();
FFiniteBoundaries_LReal();
FRelations_Real();
FRelations_LReal();
FNonFinite_Real();
FNonFinite_LReal();

FClassification_Real();
FArrayClassification_Real();
FClassification_LReal();
FArrayClassification_LReal();
END_METHOD

END_FUNCTION_BLOCK

// ---- SelfTests/TestCases/TestSuite_AssertionFloatingPoint/Test_AssertionTolerance_Real.TcPOU
{region 'Documentation'}
(*!
<summary>Checks REAL absolute tolerance boundaries and Error escalation in both relations.</summary>
<description>
Named rows separate independent comparisons by a disabled reset call.
Only explicitly marked escalation rows retain the preceding subject result.
Outer Assertions latch every observation before advancing to the next row.
All finite comparison values are exact binary fractions; expected results are literal.
ErrorAfterEqualFailure and ErrorAfterNotEqualFailure exercise each held-Failed guard.
RepeatedError and ValidInputsAfterError require held Error without another finding.
Intentional findings remain in the local capture; no production algorithm is copied.
</description>
*)
{endregion}
FUNCTION_BLOCK Test_AssertionTolerance_Real EXTENDS TestCaseBase
VAR
    FEqualSubject : AssertEqualTolerance_Real;
    FNotEqualSubject : AssertNotEqualTolerance_Real;
    FActual : REAL;
    FExpected : REAL;
    FTolerance : REAL;
    FExpectedEqualResult : E_Result;
    FExpectedNotEqualResult : E_Result;
    FExpectedFindings : UDINT;
    FExpectedEqualFinding : E_Result;
    FExpectedNotEqualFinding : E_Result;
    FCapture : EventBuffer;
    FEvents : ARRAY[1..CaptureLength] OF ST_Event;
    FCaptureFifo : ST_FifoStatus;
    FCaptureStatus : ST_EventBufferStatus;
    FRow : UINT;
    FRowPrepared : BOOL;
    FPreserveResults : BOOL;
    FObservationReady : BOOL;
    FChecked : BOOL;
    FSetupValid : BOOL;
END_VAR
VAR
    FEqualResult : AssertTrue;
    FEqualResultMatches : BOOL;
    FNotEqualResult : AssertTrue;
    FNotEqualResultMatches : BOOL;
    FCaptureIntegrity : AssertTrue;
    FCaptureIntegrityMatches : BOOL;
    FFindingDetails : AssertTrue;
    FFindingDetailsMatch : BOOL;
END_VAR
VAR CONSTANT
    CaptureLength : UINT := 8;
    EqualValues : UINT := 1;
    InsideLower : UINT := 2;
    InsideUpper : UINT := 3;
    AtLowerBoundary : UINT := 4;
    AtUpperBoundary : UINT := 5;
    OutsideLower : UINT := 6;
    OutsideUpper : UINT := 7;
    ZeroToleranceEqual : UINT := 8;
    ZeroToleranceDifferent : UINT := 9;
    NegativeTolerance : UINT := 10;
    EqualFailureBeforeError : UINT := 11;
    ErrorAfterEqualFailure : UINT := 12;
    RepeatedError : UINT := 13;
    ValidInputsAfterError : UINT := 14;
    NotEqualFailureBeforeError : UINT := 15;
    ErrorAfterNotEqualFailure : UINT := 16;
    ResetRestoresEvaluation : UINT := 17;
    LastRow : UINT := ResetRestoresEvaluation;
END_VAR

SUPER^();

{region 'Documentation'}
(*!
<summary>Collects only outer checking Assertions, never intentional subject findings.</summary>
*)
{endregion}
METHOD PROTECTED AggregateResults
VAR_INPUT
    Aggregator : I_ResultAggregator; //! Borrowed result sink owned by the outer Test Case; add this test's checking Assertions without resetting or retaining the sink.
END_VAR
Aggregator.AddProvider(Provider := FEqualResult);
Aggregator.AddProvider(Provider := FNotEqualResult);
Aggregator.AddProvider(Provider := FCaptureIntegrity);
Aggregator.AddProvider(Provider := FFindingDetails);
END_METHOD

{region 'Documentation'}
(*!
<summary>Calls each inherited production Assertion once using the selected row.</summary>
*)
{endregion}
METHOD PRIVATE CallSubjects
VAR_INPUT
    Enable : BOOL; //! Observation-enable input forwarded to the controlled Assertion subjects for this call.
END_VAR
FEqualSubject(Enable := Enable,
    State := E_State.Running,
    IN := FActual,
    Expected := FExpected,
    Tolerance := FTolerance);
FNotEqualSubject(Enable := Enable,
    State := E_State.Running,
    IN := FActual,
    Expected := FExpected,
    Tolerance := FTolerance);
END_METHOD

{region 'Documentation'}
(*!
<summary>Extends base validation with subject and checking-Assertion setup.</summary>
*)
{endregion}
METHOD PROTECTED CheckInitialization : BOOL //! TRUE when the inherited initialization check and this concrete fixture check both accept the setup.
CheckInitialization := SUPER^.CheckInitialization();
IF NOT CheckInitialization THEN
    RETURN;
END_IF;

